   #"Output Barcode" := ("Expected/Value_All".V = "Expected/Value_All".Expected_1) OR ("Expected/Value_All".V = "Expected/Value_All".Expected_2) OR ("Expected/Value_All".V = "Expected/Value_All".Expected_3) OR ("Expected/Value_All".V = "Expected/Value_All".Expected_4) OR ("Expected/Value_All".V = "Expected/Value_All".Expected_5) OR ("Expected/Value_All".V = "Expected/Value_All".Expected_6) OR ("Expected/Value_All".V = "Expected/Value_All".Expected_7) OR ("Expected/Value_All".V = "Expected/Value_All".Expected_8) OR ("Expected/Value_All".V = "Expected/Value_All".Expected_9) OR ("Expected/Value_All".V = "Expected/Value_All".Expected_10) OR ("Expected/Value_All".V = "Expected/Value_All".Expected_11) OR ("Expected/Value_All".V = "Expected/Value_All".Expected_12) OR ("Expected/Value_All".V = "Expected/Value_All".Expected_13) OR ("Expected/Value_All".V = "Expected/Value_All".Expected_14) OR ("Expected/Value_All".V = "Expected/Value_All".Expected_15) OR ("Expected/Value_All".V = "Expected/Value_All".Expected_16) OR ("Expected/Value_All".V = "Expected/Value_All".Expected_17) OR ("Expected/Value_All".V = "Expected/Value_All".Expected_18) OR ("Expected/Value_All".V = "Expected/Value_All".Expected_19) OR ("Expected/Value_All".V = "Expected/Value_All".Expected_20) OR ("Expected/Value_All".V = "Expected/Value_All".Expected_21) OR ("Expected/Value_All".V = "Expected/Value_All".Expected_22) OR ("Expected/Value_All".V = "Expected/Value_All".Expected_23) OR ("Expected/Value_All".V = "Expected/Value_All".Expected_24) OR ("Expected/Value_All".V = "Expected/Value_All".Expected_25) OR ("Expected/Value_All".V = "Expected/Value_All".Expected_26) OR ("Expected/Value_All".V = "Expected/Value_All".Expected_27) OR ("Expected/Value_All".V = "Expected/Value_All".Expected_28) OR ("Expected/Value_All".V = "Expected/Value_All".Expected_29) OR ("Expected/Value_All".V = "Expected/Value_All".Expected_30) OR ("Expected/Value_All".V = "Expected/Value_All".Expected_31) OR ("Expected/Value_All".V = "Expected/Value_All".Expected_32) OR ("Expected/Value_All".V = "Expected/Value_All".Expected_33) OR ("Expected/Value_All".V = "Expected/Value_All".Expected_34) OR ("Expected/Value_All".V = "Expected/Value_All".Expected_35) OR ("Expected/Value_All".V = "Expected/Value_All".Expected_36) OR ("Expected/Value_All".V = "Expected/Value_All".Expected_37) OR ("Expected/Value_All".V = "Expected/Value_All".Expected_38) OR ("Expected/Value_All".V = "Expected/Value_All".Expected_39) OR ("Expected/Value_All".V = "Expected/Value_All".Expected_40) OR ("Expected/Value_All".V = "Expected/Value_All".Expected_41) OR ("Expected/Value_All".V = "Expected/Value_All".Expected_42) OR ("Expected/Value_All".V = "Expected/Value_All".Expected_43) OR ("Expected/Value_All".V = "Expected/Value_All".Expected_44) OR ("Expected/Value_All".V = "Expected/Value_All".Expected_45) OR ("Expected/Value_All".V = "Expected/Value_All".Expected_46) OR ("Expected/Value_All".V = "Expected/Value_All".Expected_47) OR ("Expected/Value_All".V = "Expected/Value_All".Expected_48) OR ("Expected/Value_All".V = "Expected/Value_All".Expected_49) OR ("Expected/Value_All".V = "Expected/Value_All".Expected_50) OR ("Expected/Value_All".V = "Expected/Value_All".Expected_51) OR ("Expected/Value_All".V = "Expected/Value_All".Expected_52) OR ("Expected/Value_All".V = "Expected/Value_All".Expected_53) OR ("Expected/Value_All".V = "Expected/Value_All".Expected_54) OR ("Expected/Value_All".V = "Expected/Value_All".Expected_55) OR ("Expected/Value_All".V = "Expected/Value_All".Expected_56) OR ("Expected/Value_All".V = "Expected/Value_All".Expected_57) OR ("Expected/Value_All".V = "Expected/Value_All".Expected_58) OR ("Expected/Value_All".V = "Expected/Value_All".Expected_59) OR ("Expected/Value_All".V = "Expected/Value_All".Expected_60) OR ("Expected/Value_All".V = "Expected/Value_All".Expected_61) OR ("Expected/Value_All".V = "Expected/Value_All".Expected_62) OR ("Expected/Value_All".V = "Expected/Value_All".Expected_63) OR ("Expected/Value_All".V = "Expected/Value_All".Expected_64) OR ("Expected/Value_All".V = "Expected/Value_All".Expected_65) OR ("Expected/Value_All".V = "Expected/Value_All".Expected_66) OR ("Expected/Value_All".V = "Expected/Value_All".Expected_67) OR ("Expected/Value_All".V = "Expected/Value_All".Expected_68) OR ("Expected/Value_All".V = "Expected/Value_All".Expected_69) OR ("Expected/Value_All".V = "Expected/Value_All".Expected_70) OR ("Expected/Value_All".V = "Expected/Value_All".Expected_71) OR ("Expected/Value_All".V = "Expected/Value_All".Expected_72) OR ("Expected/Value_All".V = "Expected/Value_All".Expected_73) OR ("Expected/Value_All".V = "Expected/Value_All".Expected_74) OR ("Expected/Value_All".V = "Expected/Value_All".Expected_75) OR ("Expected/Value_All".V = "Expected/Value_All".Expected_76) OR ("Expected/Value_All".V = "Expected/Value_All".Expected_77) OR ("Expected/Value_All".V = "Expected/Value_All".Expected_78) OR ("Expected/Value_All".V = "Expected/Value_All".Expected_79) OR ("Expected/Value_All".V = "Expected/Value_All".Expected_80) OR ("Expected/Value_All".V = "Expected/Value_All".Expected_81) OR ("Expected/Value_All".V = "Expected/Value_All".Expected_82) OR ("Expected/Value_All".V = "Expected/Value_All".Expected_83) OR ("Expected/Value_All".V = "Expected/Value_All".Expected_84) OR ("Expected/Value_All".V = "Expected/Value_All".Expected_85) OR ("Expected/Value_All".V = "Expected/Value_All".Expected_86) OR ("Expected/Value_All".V = "Expected/Value_All".Expected_87) OR ("Expected/Value_All".V = "Expected/Value_All".Expected_88) OR ("Expected/Value_All".V = "Expected/Value_All".Expected_89) OR ("Expected/Value_All".V = "Expected/Value_All".Expected_90) OR ("Expected/Value_All".V = "Expected/Value_All".Expected_91) OR ("Expected/Value_All".V = "Expected/Value_All".Expected_92) OR ("Expected/Value_All".V = "Expected/Value_All".Expected_93) OR ("Expected/Value_All".V = "Expected/Value_All".Expected_94) OR ("Expected/Value_All".V = "Expected/Value_All".Expected_95) OR ("Expected/Value_All".V = "Expected/Value_All".Expected_96) OR ("Expected/Value_All".V = "Expected/Value_All".Expected_97) OR ("Expected/Value_All".V = "Expected/Value_All".Expected_98) OR ("Expected/Value_All".V = "Expected/Value_All".Expected_99) OR ("Expected/Value_All".V = "Expected/Value_All".Expected_100) OR ("Expected/Value_All".V = "Expected/Value_All".Expected_101) OR ("Expected/Value_All".V = "Expected/Value_All".Expected_102) OR ("Expected/Value_All".V = "Expected/Value_All".Expected_103) OR ("Expected/Value_All".V = "Expected/Value_All".Expected_104) OR ("Expected/Value_All".V = "Expected/Value_All".Expected_105) OR ("Expected/Value_All".V = "Expected/Value_All".Expected_106) OR ("Expected/Value_All".V = "Expected/Value_All".Expected_107) OR ("Expected/Value_All".V = "Expected/Value_All".Expected_108) OR ("Expected/Value_All".V = "Expected/Value_All".Expected_109) OR ("Expected/Value_All".V = "Expected/Value_All".Expected_110) OR ("Expected/Value_All".V = "Expected/Value_All".Expected_111) OR ("Expected/Value_All".V = "Expected/Value_All".Expected_112) OR ("Expected/Value_All".V = "Expected/Value_All".Expected_113) OR ("Expected/Value_All".V = "Expected/Value_All".Expected_114) OR ("Expected/Value_All".V = "Expected/Value_All".Expected_115) OR ("Expected/Value_All".V = "Expected/Value_All".Expected_116) OR ("Expected/Value_All".V = "Expected/Value_All".Expected_117) OR ("Expected/Value_All".V = "Expected/Value_All".Expected_118) OR ("Expected/Value_All".V = "Expected/Value_All".Expected_119) OR ("Expected/Value_All".V = "Expected/Value_All".Expected_120) OR ("Expected/Value_All".V = "Expected/Value_All".Expected_121) OR ("Expected/Value_All".V = "Expected/Value_All".Expected_122) OR ("Expected/Value_All".V = "Expected/Value_All".Expected_123) OR ("Expected/Value_All".V = "Expected/Value_All".Expected_124) OR ("Expected/Value_All".V = "Expected/Value_All".Expected_125) OR ("Expected/Value_All".V = "Expected/Value_All".Expected_126) OR ("Expected/Value_All".V = "Expected/Value_All".Expected_127) OR ("Expected/Value_All".V = "Expected/Value_All".Expected_128) OR ("Expected/Value_All".V = "Expected/Value_All".Expected_129) OR ("Expected/Value_All".V = "Expected/Value_All".Expected_130) OR ("Expected/Value_All".V = "Expected/Value_All".Expected_131) OR ("Expected/Value_All".V = "Expected/Value_All".Expected_132) OR ("Expected/Value_All".V = "Expected/Value_All".Expected_133) OR ("Expected/Value_All".V = "Expected/Value_All".Expected_134) OR ("Expected/Value_All".V = "Expected/Value_All".Expected_135) OR ("Expected/Value_All".V = "Expected/Value_All".Expected_136) OR ("Expected/Value_All".V = "Expected/Value_All".Expected_137) OR ("Expected/Value_All".V = "Expected/Value_All".Expected_138) OR ("Expected/Value_All".V = "Expected/Value_All".Expected_139) OR ("Expected/Value_All".V = "Expected/Value_All".Expected_140) OR ("Expected/Value_All".V = "Expected/Value_All".Expected_141) OR ("Expected/Value_All".V = "Expected/Value_All".Expected_142) OR ("Expected/Value_All".V = "Expected/Value_All".Expected_143) OR ("Expected/Value_All".V = "Expected/Value_All".Expected_144) OR ("Expected/Value_All".V = "Expected/Value_All".Expected_145) OR ("Expected/Value_All".V = "Expected/Value_All".Expected_146) OR ("Expected/Value_All".V = "Expected/Value_All".Expected_147) OR ("Expected/Value_All".V = "Expected/Value_All".Expected_148) OR ("Expected/Value_All".V = "Expected/Value_All".Expected_149) OR ("Expected/Value_All".V = "Expected/Value_All".Expected_150) OR ("Expected/Value_All".V = "Expected/Value_All".Expected_151) OR ("Expected/Value_All".V = "Expected/Value_All".Expected_152) OR ("Expected/Value_All".V = "Expected/Value_All".Expected_153) OR ("Expected/Value_All".V = "Expected/Value_All".Expected_154) OR ("Expected/Value_All".V = "Expected/Value_All".Expected_155) OR ("Expected/Value_All".V = "Expected/Value_All".Expected_156) OR ("Expected/Value_All".V = "Expected/Value_All".Expected_157) OR ("Expected/Value_All".V = "Expected/Value_All".Expected_158) OR ("Expected/Value_All".V = "Expected/Value_All".Expected_159) OR ("Expected/Value_All".V = "Expected/Value_All".Expected_160) OR ("Expected/Value_All".V = "Expected/Value_All".Expected_161) OR ("Expected/Value_All".V = "Expected/Value_All".Expected_162) OR ("Expected/Value_All".V = "Expected/Value_All".Expected_163) OR ("Expected/Value_All".V = "Expected/Value_All".Expected_164) OR ("Expected/Value_All".V = "Expected/Value_All".Expected_165) OR ("Expected/Value_All".V = "Expected/Value_All".Expected_166) OR ("Expected/Value_All".V = "Expected/Value_All".Expected_167) OR ("Expected/Value_All".V = "Expected/Value_All".Expected_168) OR ("Expected/Value_All".V = "Expected/Value_All".Expected_169) OR ("Expected/Value_All".V = "Expected/Value_All".Expected_170) OR ("Expected/Value_All".V = "Expected/Value_All".Expected_171) OR ("Expected/Value_All".V = "Expected/Value_All".Expected_172) OR ("Expected/Value_All".V = "Expected/Value_All".Expected_173) OR ("Expected/Value_All".V = "Expected/Value_All".Expected_174) OR ("Expected/Value_All".V = "Expected/Value_All".Expected_175) OR ("Expected/Value_All".V = "Expected/Value_All".Expected_176) OR ("Expected/Value_All".V = "Expected/Value_All".Expected_177) OR ("Expected/Value_All".V = "Expected/Value_All".Expected_178) OR ("Expected/Value_All".V = "Expected/Value_All".Expected_179) OR ("Expected/Value_All".V = "Expected/Value_All".Expected_180) OR ("Expected/Value_All".V = "Expected/Value_All".Expected_181) OR ("Expected/Value_All".V = "Expected/Value_All".Expected_182) OR ("Expected/Value_All".V = "Expected/Value_All".Expected_183) OR ("Expected/Value_All".V = "Expected/Value_All".Expected_184) OR ("Expected/Value_All".V = "Expected/Value_All".Expected_185) OR ("Expected/Value_All".V = "Expected/Value_All".Expected_186) OR ("Expected/Value_All".V = "Expected/Value_All".Expected_187) OR ("Expected/Value_All".V = "Expected/Value_All".Expected_188) OR ("Expected/Value_All".V = "Expected/Value_All".Expected_189) OR ("Expected/Value_All".V = "Expected/Value_All".Expected_190) OR ("Expected/Value_All".V = "Expected/Value_All".Expected_191) OR ("Expected/Value_All".V = "Expected/Value_All".Expected_192) OR ("Expected/Value_All".V = "Expected/Value_All".Expected_193) OR ("Expected/Value_All".V = "Expected/Value_All".Expected_194) OR ("Expected/Value_All".V = "Expected/Value_All".Expected_195) OR ("Expected/Value_All".V = "Expected/Value_All".Expected_196) OR ("Expected/Value_All".V = "Expected/Value_All".Expected_197) OR ("Expected/Value_All".V = "Expected/Value_All".Expected_198) OR ("Expected/Value_All".V = "Expected/Value_All".Expected_199) OR ("Expected/Value_All".V = "Expected/Value_All".Expected_200) OR ("Expected/Value_All".V = "Expected/Value_All".Expected_201) OR ("Expected/Value_All".V = "Expected/Value_All".Expected_202) OR ("Expected/Value_All".V = "Expected/Value_All".Expected_203) OR ("Expected/Value_All".V = "Expected/Value_All".Expected_204) OR ("Expected/Value_All".V = "Expected/Value_All".Expected_205) OR ("Expected/Value_All".V = "Expected/Value_All".Expected_206) OR ("Expected/Value_All".V = "Expected/Value_All".Expected_207) OR ("Expected/Value_All".V = "Expected/Value_All".Expected_208) OR ("Expected/Value_All".V = "Expected/Value_All".Expected_209) OR ("Expected/Value_All".V = "Expected/Value_All".Expected_210) OR ("Expected/Value_All".V = "Expected/Value_All".Expected_211) OR ("Expected/Value_All".V = "Expected/Value_All".Expected_212) OR ("Expected/Value_All".V = "Expected/Value_All".Expected_213) OR ("Expected/Value_All".V = "Expected/Value_All".Expected_214) OR ("Expected/Value_All".V = "Expected/Value_All".Expected_215) OR ("Expected/Value_All".V = "Expected/Value_All".Expected_216) OR ("Expected/Value_All".V = "Expected/Value_All".Expected_217) OR ("Expected/Value_All".V = "Expected/Value_All".Expected_218) OR ("Expected/Value_All".V = "Expected/Value_All".Expected_219) OR ("Expected/Value_All".V = "Expected/Value_All".Expected_220) OR ("Expected/Value_All".V = "Expected/Value_All".Expected_221) OR ("Expected/Value_All".V = "Expected/Value_All".Expected_222) OR ("Expected/Value_All".V = "Expected/Value_All".Expected_223) OR ("Expected/Value_All".V = "Expected/Value_All".Expected_224) OR ("Expected/Value_All".V = "Expected/Value_All".Expected_225) OR ("Expected/Value_All".V = "Expected/Value_All".Expected_226) OR ("Expected/Value_All".V = "Expected/Value_All".Expected_227) OR ("Expected/Value_All".V = "Expected/Value_All".Expected_228) OR ("Expected/Value_All".V = "Expected/Value_All".Expected_229) OR ("Expected/Value_All".V = "Expected/Value_All".Expected_230) OR ("Expected/Value_All".V = "Expected/Value_All".Expected_231) OR ("Expected/Value_All".V = "Expected/Value_All".Expected_232) OR ("Expected/Value_All".V = "Expected/Value_All".Expected_233) OR ("Expected/Value_All".V = "Expected/Value_All".Expected_234) OR ("Expected/Value_All".V = "Expected/Value_All".Expected_235) OR ("Expected/Value_All".V = "Expected/Value_All".Expected_236) OR ("Expected/Value_All".V = "Expected/Value_All".Expected_237) OR ("Expected/Value_All".V = "Expected/Value_All".Expected_238) OR ("Expected/Value_All".V = "Expected/Value_All".Expected_239) OR ("Expected/Value_All".V = "Expected/Value_All".Expected_240) OR ("Expected/Value_All".V = "Expected/Value_All".Expected_241) OR ("Expected/Value_All".V = "Expected/Value_All".Expected_242) OR ("Expected/Value_All".V = "Expected/Value_All".Expected_243) OR ("Expected/Value_All".V = "Expected/Value_All".Expected_244) OR ("Expected/Value_All".V = "Expected/Value_All".Expected_245) OR ("Expected/Value_All".V = "Expected/Value_All".Expected_246) OR ("Expected/Value_All".V = "Expected/Value_All".Expected_247) OR ("Expected/Value_All".V = "Expected/Value_All".Expected_248) OR ("Expected/Value_All".V = "Expected/Value_All".Expected_249) OR ("Expected/Value_All".V = "Expected/Value_All".Expected_250) OR ("Expected/Value_All".V = "Expected/Value_All".Expected_251) OR ("Expected/Value_All".V = "Expected/Value_All".Expected_252) OR ("Expected/Value_All".V = "Expected/Value_All".Expected_253) OR ("Expected/Value_All".V = "Expected/Value_All".Expected_254) OR ("Expected/Value_All".V = "Expected/Value_All".Expected_255) OR ("Expected/Value_All".V = "Expected/Value_All".Expected_256) OR ("Expected/Value_All".V = "Expected/Value_All".Expected_257) OR ("Expected/Value_All".V = "Expected/Value_All".Expected_258) OR ("Expected/Value_All".V = "Expected/Value_All".Expected_259) OR ("Expected/Value_All".V = "Expected/Value_All".Expected_260) OR ("Expected/Value_All".V = "Expected/Value_All".Expected_261) OR ("Expected/Value_All".V = "Expected/Value_All".Expected_262) OR ("Expected/Value_All".V = "Expected/Value_All".Expected_263) OR ("Expected/Value_All".V = "Expected/Value_All".Expected_264) OR ("Expected/Value_All".V = "Expected/Value_All".Expected_265) OR ("Expected/Value_All".V = "Expected/Value_All".Expected_266) OR ("Expected/Value_All".V = "Expected/Value_All".Expected_267) OR ("Expected/Value_All".V = "Expected/Value_All".Expected_268) OR ("Expected/Value_All".V = "Expected/Value_All".Expected_269) OR ("Expected/Value_All".V = "Expected/Value_All".Expected_270) OR ("Expected/Value_All".V = "Expected/Value_All".Expected_271) OR ("Expected/Value_All".V = "Expected/Value_All".Expected_272) OR ("Expected/Value_All".V = "Expected/Value_All".Expected_273) OR ("Expected/Value_All".V = "Expected/Value_All".Expected_274) OR ("Expected/Value_All".V = "Expected/Value_All".Expected_275) OR ("Expected/Value_All".V = "Expected/Value_All".Expected_276) OR ("Expected/Value_All".V = "Expected/Value_All".Expected_277) OR ("Expected/Value_All".V = "Expected/Value_All".Expected_278) OR ("Expected/Value_All".V = "Expected/Value_All".Expected_279) OR ("Expected/Value_All".V = "Expected/Value_All".Expected_280) OR ("Expected/Value_All".V = "Expected/Value_All".Expected_281) OR ("Expected/Value_All".V = "Expected/Value_All".Expected_282) OR ("Expected/Value_All".V = "Expected/Value_All".Expected_283) OR ("Expected/Value_All".V = "Expected/Value_All".Expected_284) OR ("Expected/Value_All".V = "Expected/Value_All".Expected_285) OR ("Expected/Value_All".V = "Expected/Value_All".Expected_286) OR ("Expected/Value_All".V = "Expected/Value_All".Expected_287) OR ("Expected/Value_All".V = "Expected/Value_All".Expected_288) OR ("Expected/Value_All".V = "Expected/Value_All".Expected_289) OR ("Expected/Value_All".V = "Expected/Value_All".Expected_290) OR ("Expected/Value_All".V = "Expected/Value_All".Expected_291) OR ("Expected/Value_All".V = "Expected/Value_All".Expected_292) OR ("Expected/Value_All".V = "Expected/Value_All".Expected_293) OR ("Expected/Value_All".V = "Expected/Value_All".Expected_294) OR ("Expected/Value_All".V = "Expected/Value_All".Expected_295) OR ("Expected/Value_All".V = "Expected/Value_All".Expected_296) OR ("Expected/Value_All".V = "Expected/Value_All".Expected_297) OR ("Expected/Value_All".V = "Expected/Value_All".Expected_298) OR ("Expected/Value_All".V = "Expected/Value_All".Expected_299) OR ("Expected/Value_All".V = "Expected/Value_All".Expected_300) OR ("Expected/Value_All".V = "Expected/Value_All".Expected_301) OR ("Expected/Value_All".V = "Expected/Value_All".Expected_302) OR ("Expected/Value_All".V = "Expected/Value_All".Expected_303) OR ("Expected/Value_All".V = "Expected/Value_All".Expected_304) OR ("Expected/Value_All".V = "Expected/Value_All".Expected_305) OR ("Expected/Value_All".V = "Expected/Value_All".Expected_306) OR ("Expected/Value_All".V = "Expected/Value_All".Expected_307) OR ("Expected/Value_All".V = "Expected/Value_All".Expected_308) OR ("Expected/Value_All".V = "Expected/Value_All".Expected_309) OR ("Expected/Value_All".V = "Expected/Value_All".Expected_310) OR ("Expected/Value_All".V = "Expected/Value_All".Expected_311) OR ("Expected/Value_All".V = "Expected/Value_All".Expected_312) OR ("Expected/Value_All".V = "Expected/Value_All".Expected_313) OR ("Expected/Value_All".V = "Expected/Value_All".Expected_314) OR ("Expected/Value_All".V = "Expected/Value_All".Expected_315) OR ("Expected/Value_All".V = "Expected/Value_All".Expected_316) OR ("Expected/Value_All".V = "Expected/Value_All".Expected_317) OR ("Expected/Value_All".V = "Expected/Value_All".Expected_318) OR ("Expected/Value_All".V = "Expected/Value_All".Expected_319) OR ("Expected/Value_All".V = "Expected/Value_All".Expected_320) OR ("Expected/Value_All".V = "Expected/Value_All".Expected_321) OR ("Expected/Value_All".V = "Expected/Value_All".Expected_322) OR ("Expected/Value_All".V = "Expected/Value_All".Expected_323) OR ("Expected/Value_All".V = "Expected/Value_All".Expected_324) OR ("Expected/Value_All".V = "Expected/Value_All".Expected_325) OR ("Expected/Value_All".V = "Expected/Value_All".Expected_326) OR ("Expected/Value_All".V = "Expected/Value_All".Expected_327) OR ("Expected/Value_All".V = "Expected/Value_All".Expected_328) OR ("Expected/Value_All".V = "Expected/Value_All".Expected_329) OR ("Expected/Value_All".V = "Expected/Value_All".Expected_330) OR ("Expected/Value_All".V = "Expected/Value_All".Expected_331) OR ("Expected/Value_All".V = "Expected/Value_All".Expected_332) OR ("Expected/Value_All".V = "Expected/Value_All".Expected_333) OR ("Expected/Value_All".V = "Expected/Value_All".Expected_334) OR ("Expected/Value_All".V = "Expected/Value_All".Expected_335) OR ("Expected/Value_All".V = "Expected/Value_All".Expected_336) OR ("Expected/Value_All".V = "Expected/Value_All".Expected_337) OR ("Expected/Value_All".V = "Expected/Value_All".Expected_338) OR ("Expected/Value_All".V = "Expected/Value_All".Expected_339) OR ("Expected/Value_All".V = "Expected/Value_All".Expected_340) OR ("Expected/Value_All".V = "Expected/Value_All".Expected_341) OR ("Expected/Value_All".V = "Expected/Value_All".Expected_342) OR ("Expected/Value_All".V = "Expected/Value_All".Expected_343) OR ("Expected/Value_All".V = "Expected/Value_All".Expected_344) OR ("Expected/Value_All".V = "Expected/Value_All".Expected_345) OR ("Expected/Value_All".V = "Expected/Value_All".Expected_346) OR ("Expected/Value_All".V = "Expected/Value_All".Expected_347) OR ("Expected/Value_All".V = "Expected/Value_All".Expected_348) OR ("Expected/Value_All".V = "Expected/Value_All".Expected_349) OR ("Expected/Value_All".V = "Expected/Value_All".Expected_350) OR ("Expected/Value_All".V = "Expected/Value_All".Expected_351) OR ("Expected/Value_All".V = "Expected/Value_All".Expected_352) OR ("Expected/Value_All".V = "Expected/Value_All".Expected_353) OR ("Expected/Value_All".V = "Expected/Value_All".Expected_354) OR ("Expected/Value_All".V = "Expected/Value_All".Expected_355) OR ("Expected/Value_All".V = "Expected/Value_All".Expected_356) OR ("Expected/Value_All".V = "Expected/Value_All".Expected_357) OR ("Expected/Value_All".V = "Expected/Value_All".Expected_358) OR ("Expected/Value_All".V = "Expected/Value_All".Expected_359) OR ("Expected/Value_All".V = "Expected/Value_All".Expected_360) OR ("Expected/Value_All".V = "Expected/Value_All".Expected_361) OR ("Expected/Value_All".V = "Expected/Value_All".Expected_362) OR ("Expected/Value_All".V = "Expected/Value_All".Expected_363) OR ("Expected/Value_All".V = "Expected/Value_All".Expected_364) OR ("Expected/Value_All".V = "Expected/Value_All".Expected_365) OR ("Expected/Value_All".V = "Expected/Value_All".Expected_366) OR ("Expected/Value_All".V = "Expected/Value_All".Expected_367) OR ("Expected/Value_All".V = "Expected/Value_All".Expected_368) OR ("Expected/Value_All".V = "Expected/Value_All".Expected_369) OR ("Expected/Value_All".V = "Expected/Value_All".Expected_370) OR ("Expected/Value_All".V = "Expected/Value_All".Expected_371) OR ("Expected/Value_All".V = "Expected/Value_All".Expected_372) OR ("Expected/Value_All".V = "Expected/Value_All".Expected_373) OR ("Expected/Value_All".V = "Expected/Value_All".Expected_374) OR ("Expected/Value_All".V = "Expected/Value_All".Expected_375) OR ("Expected/Value_All".V = "Expected/Value_All".Expected_376) OR ("Expected/Value_All".V = "Expected/Value_All".Expected_377) OR ("Expected/Value_All".V = "Expected/Value_All".Expected_378) OR ("Expected/Value_All".V = "Expected/Value_All".Expected_379) OR ("Expected/Value_All".V = "Expected/Value_All".Expected_380) OR ("Expected/Value_All".V = "Expected/Value_All".Expected_381) OR ("Expected/Value_All".V = "Expected/Value_All".Expected_382) OR ("Expected/Value_All".V = "Expected/Value_All".Expected_383) OR ("Expected/Value_All".V = "Expected/Value_All".Expected_384) OR ("Expected/Value_All".V = "Expected/Value_All".Expected_385) OR ("Expected/Value_All".V = "Expected/Value_All".Expected_386) OR ("Expected/Value_All".V = "Expected/Value_All".Expected_387) OR ("Expected/Value_All".V = "Expected/Value_All".Expected_388) OR ("Expected/Value_All".V = "Expected/Value_All".Expected_389) OR ("Expected/Value_All".V = "Expected/Value_All".Expected_390) OR ("Expected/Value_All".V = "Expected/Value_All".Expected_391) OR ("Expected/Value_All".V = "Expected/Value_All".Expected_392) OR ("Expected/Value_All".V = "Expected/Value_All".Expected_393) OR ("Expected/Value_All".V = "Expected/Value_All".Expected_394) OR ("Expected/Value_All".V = "Expected/Value_All".Expected_395) OR ("Expected/Value_All".V = "Expected/Value_All".Expected_396) OR ("Expected/Value_All".V = "Expected/Value_All".Expected_397) OR ("Expected/Value_All".V = "Expected/Value_All".Expected_398) OR ("Expected/Value_All".V = "Expected/Value_All".Expected_399) OR ("Expected/Value_All".V = "Expected/Value_All".Expected_400) OR ("Expected/Value_All".V = "Expected/Value_All".Expected_401) OR ("Expected/Value_All".V = "Expected/Value_All".Expected_402) OR ("Expected/Value_All".V = "Expected/Value_All".Expected_403) OR ("Expected/Value_All".V = "Expected/Value_All".Expected_404) OR ("Expected/Value_All".V = "Expected/Value_All".Expected_405) OR ("Expected/Value_All".V = "Expected/Value_All".Expected_406) OR ("Expected/Value_All".V = "Expected/Value_All".Expected_407) OR ("Expected/Value_All".V = "Expected/Value_All".Expected_408) OR ("Expected/Value_All".V = "Expected/Value_All".Expected_409) OR ("Expected/Value_All".V = "Expected/Value_All".Expected_410) OR ("Expected/Value_All".V = "Expected/Value_All".Expected_411) OR ("Expected/Value_All".V = "Expected/Value_All".Expected_412) OR ("Expected/Value_All".V = "Expected/Value_All".Expected_413) OR ("Expected/Value_All".V = "Expected/Value_All".Expected_414) OR ("Expected/Value_All".V = "Expected/Value_All".Expected_415) OR ("Expected/Value_All".V = "Expected/Value_All".Expected_416) OR ("Expected/Value_All".V = "Expected/Value_All".Expected_417) OR ("Expected/Value_All".V = "Expected/Value_All".Expected_418) OR ("Expected/Value_All".V = "Expected/Value_All".Expected_419) OR ("Expected/Value_All".V = "Expected/Value_All".Expected_420) OR ("Expected/Value_All".V = "Expected/Value_All".Expected_421) OR ("Expected/Value_All".V = "Expected/Value_All".Expected_422) OR ("Expected/Value_All".V = "Expected/Value_All".Expected_423) OR ("Expected/Value_All".V = "Expected/Value_All".Expected_424) OR ("Expected/Value_All".V = "Expected/Value_All".Expected_425) OR ("Expected/Value_All".V = "Expected/Value_All".Expected_426) OR ("Expected/Value_All".V = "Expected/Value_All".Expected_427) OR ("Expected/Value_All".V = "Expected/Value_All".Expected_428) OR ("Expected/Value_All".V = "Expected/Value_All".Expected_429) OR ("Expected/Value_All".V = "Expected/Value_All".Expected_430) OR ("Expected/Value_All".V = "Expected/Value_All".Expected_431) OR ("Expected/Value_All".V = "Expected/Value_All".Expected_432) OR ("Expected/Value_All".V = "Expected/Value_All".Expected_433) OR ("Expected/Value_All".V = "Expected/Value_All".Expected_434) OR ("Expected/Value_All".V = "Expected/Value_All".Expected_435) OR ("Expected/Value_All".V = "Expected/Value_All".Expected_436) OR ("Expected/Value_All".V = "Expected/Value_All".Expected_437) OR ("Expected/Value_All".V = "Expected/Value_All".Expected_438) OR ("Expected/Value_All".V = "Expected/Value_All".Expected_439) OR ("Expected/Value_All".V = "Expected/Value_All".Expected_440) OR ("Expected/Value_All".V = "Expected/Value_All".Expected_441) OR ("Expected/Value_All".V = "Expected/Value_All".Expected_442) OR ("Expected/Value_All".V = "Expected/Value_All".Expected_443) OR ("Expected/Value_All".V = "Expected/Value_All".Expected_444) OR ("Expected/Value_All".V = "Expected/Value_All".Expected_445) OR ("Expected/Value_All".V = "Expected/Value_All".Expected_446) OR ("Expected/Value_All".V = "Expected/Value_All".Expected_447) OR ("Expected/Value_All".V = "Expected/Value_All".Expected_448) OR ("Expected/Value_All".V = "Expected/Value_All".Expected_449) OR ("Expected/Value_All".V = "Expected/Value_All".Expected_450) OR ("Expected/Value_All".V = "Expected/Value_All".Expected_451) OR ("Expected/Value_All".V = "Expected/Value_All".Expected_452) OR ("Expected/Value_All".V = "Expected/Value_All".Expected_453) OR ("Expected/Value_All".V = "Expected/Value_All".Expected_454) OR ("Expected/Value_All".V = "Expected/Value_All".Expected_455) OR ("Expected/Value_All".V = "Expected/Value_All".Expected_456) OR ("Expected/Value_All".V = "Expected/Value_All".Expected_457) OR ("Expected/Value_All".V = "Expected/Value_All".Expected_458) OR ("Expected/Value_All".V = "Expected/Value_All".Expected_459) OR ("Expected/Value_All".V = "Expected/Value_All".Expected_460) OR ("Expected/Value_All".V = "Expected/Value_All".Expected_461) OR ("Expected/Value_All".V = "Expected/Value_All".Expected_462) OR ("Expected/Value_All".V = "Expected/Value_All".Expected_463) OR ("Expected/Value_All".V = "Expected/Value_All".Expected_464) OR ("Expected/Value_All".V = "Expected/Value_All".Expected_465) OR ("Expected/Value_All".V = "Expected/Value_All".Expected_466) OR ("Expected/Value_All".V = "Expected/Value_All".Expected_467) OR ("Expected/Value_All".V = "Expected/Value_All".Expected_468) OR ("Expected/Value_All".V = "Expected/Value_All".Expected_469) OR ("Expected/Value_All".V = "Expected/Value_All".Expected_470) OR ("Expected/Value_All".V = "Expected/Value_All".Expected_471) OR ("Expected/Value_All".V = "Expected/Value_All".Expected_472) OR ("Expected/Value_All".V = "Expected/Value_All".Expected_473) OR ("Expected/Value_All".V = "Expected/Value_All".Expected_474) OR ("Expected/Value_All".V = "Expected/Value_All".Expected_475) OR ("Expected/Value_All".V = "Expected/Value_All".Expected_476) OR ("Expected/Value_All".V = "Expected/Value_All".Expected_477) OR ("Expected/Value_All".V = "Expected/Value_All".Expected_478) OR ("Expected/Value_All".V = "Expected/Value_All".Expected_479) OR ("Expected/Value_All".V = "Expected/Value_All".Expected_480) OR ("Expected/Value_All".V = "Expected/Value_All".Expected_481) OR ("Expected/Value_All".V = "Expected/Value_All".Expected_482) OR ("Expected/Value_All".V = "Expected/Value_All".Expected_483) OR ("Expected/Value_All".V = "Expected/Value_All".Expected_484) OR ("Expected/Value_All".V = "Expected/Value_All".Expected_485) OR ("Expected/Value_All".V = "Expected/Value_All".Expected_486) OR ("Expected/Value_All".V = "Expected/Value_All".Expected_487) OR ("Expected/Value_All".V = "Expected/Value_All".Expected_488) OR ("Expected/Value_All".V = "Expected/Value_All".Expected_489) OR ("Expected/Value_All".V = "Expected/Value_All".Expected_490) OR ("Expected/Value_All".V = "Expected/Value_All".Expected_491) OR ("Expected/Value_All".V = "Expected/Value_All".Expected_492) OR ("Expected/Value_All".V = "Expected/Value_All".Expected_493) OR ("Expected/Value_All".V = "Expected/Value_All".Expected_494) OR ("Expected/Value_All".V = "Expected/Value_All".Expected_495) OR ("Expected/Value_All".V = "Expected/Value_All".Expected_496) OR ("Expected/Value_All".V = "Expected/Value_All".Expected_497) OR ("Expected/Value_All".V = "Expected/Value_All".Expected_498) OR ("Expected/Value_All".V = "Expected/Value_All".Expected_499) OR ("Expected/Value_All".V = "Expected/Value_All".Expected_500) OR ("Expected/Value_All".V = "Expected/Value_All".Expected_501) OR ("Expected/Value_All".V = "Expected/Value_All".Expected_502) OR ("Expected/Value_All".V = "Expected/Value_All".Expected_503) OR ("Expected/Value_All".V = "Expected/Value_All".Expected_504) OR ("Expected/Value_All".V = "Expected/Value_All".Expected_505) OR ("Expected/Value_All".V = "Expected/Value_All".Expected_506) OR ("Expected/Value_All".V = "Expected/Value_All".Expected_507) OR ("Expected/Value_All".V = "Expected/Value_All".Expected_508) OR ("Expected/Value_All".V = "Expected/Value_All".Expected_509) OR ("Expected/Value_All".V = "Expected/Value_All".Expected_510) OR ("Expected/Value_All".V = "Expected/Value_All".Expected_511) OR ("Expected/Value_All".V = "Expected/Value_All".Expected_512) OR ("Expected/Value_All".V = "Expected/Value_All".Expected_513) OR ("Expected/Value_All".V = "Expected/Value_All".Expected_514) OR ("Expected/Value_All".V = "Expected/Value_All".Expected_515) OR ("Expected/Value_All".V = "Expected/Value_All".Expected_516) OR ("Expected/Value_All".V = "Expected/Value_All".Expected_517) OR ("Expected/Value_All".V = "Expected/Value_All".Expected_518) OR ("Expected/Value_All".V = "Expected/Value_All".Expected_519) OR ("Expected/Value_All".V = "Expected/Value_All".Expected_520);
END_REGION
END_FUNCTION

FUNCTION "Expected" : Void   // FC3, LAD
{ S7_Optimized_Access := 'TRUE' }
VERSION : 0.1
   VAR_INPUT
      Expected1 : String;
      Expected2 : String;
      Expected3 : String;
      Expected4 : String;
      Expected5 : String;
      Expected6 : String;
      Expected7 : String;
      Expected8 : String;
      Expected9 : String;
      Expected10 : String;
      Expected11 : String;
      Expected12 : String;
      Expected13 : String;
      Expected14 : String;
      Expected15 : String;
      Expected16 : String;
      Expected17 : String;
      Expected18 : String;
      Expected19 : String;
      Expected20 : String;
      Expected21 : String;
      Expected22 : String;
      Expected23 : String;
      Expected24 : String;
      Expected25 : String;
      Expected26 : String;
   END_VAR
   VAR_OUTPUT
      On_Motor : Bool;
   END_VAR
BEGIN

REGION Network 1
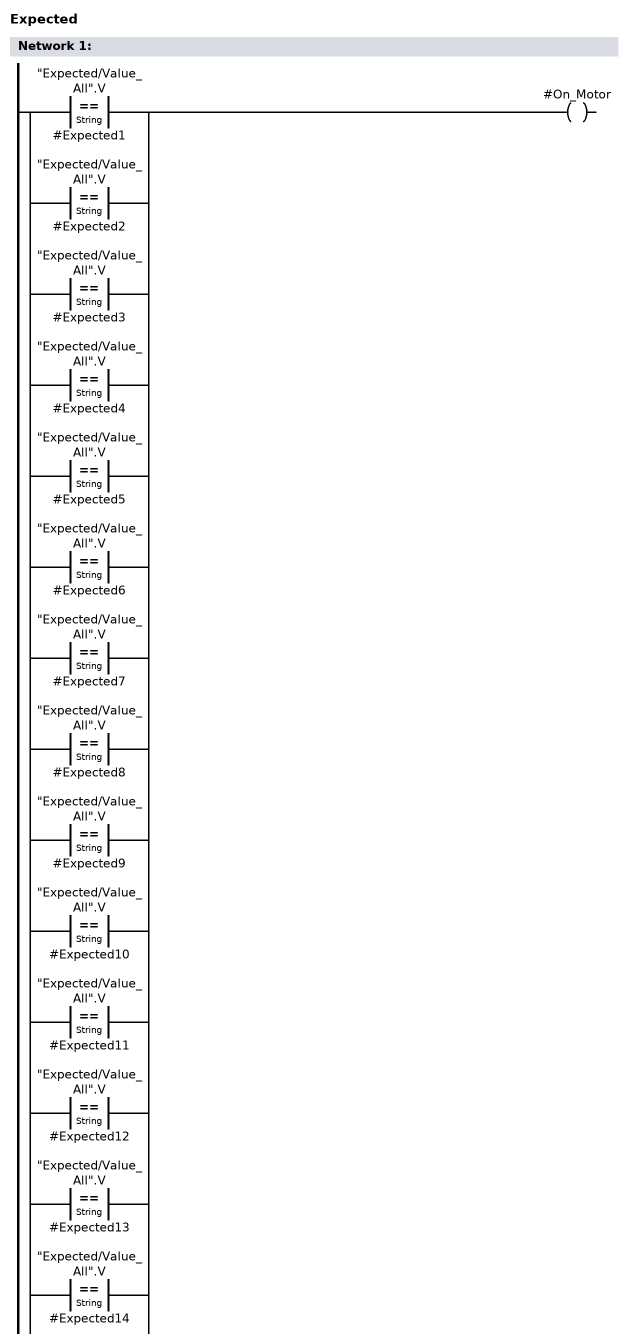
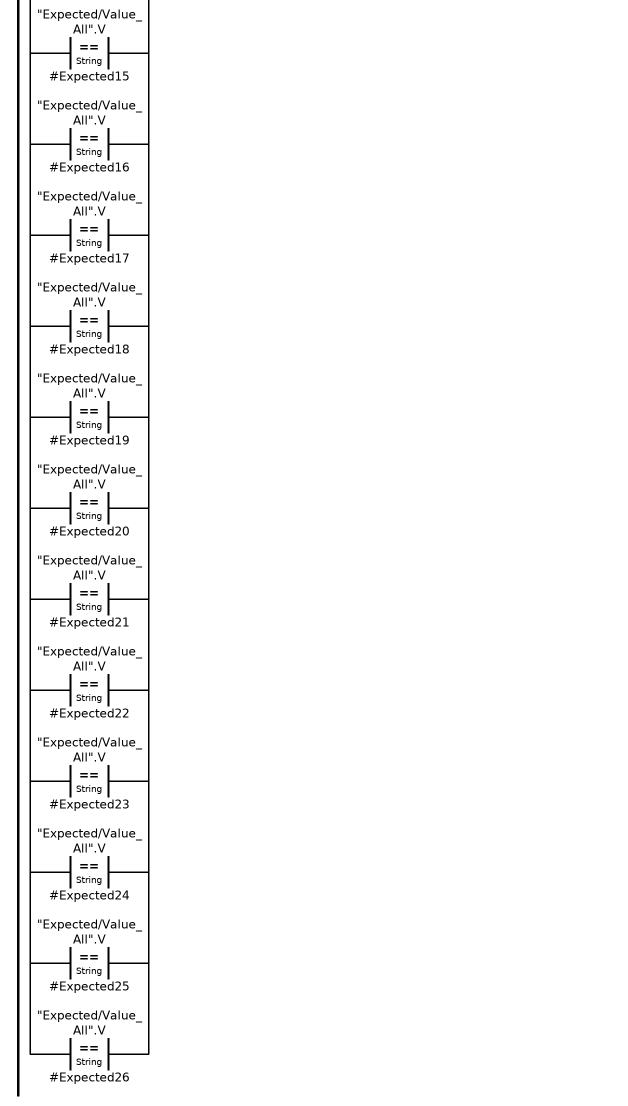
   RUNG wire#powerrail
      { S7_Templates := "SrcType := String" } EQ_Contact(in1 := "Expected/Value_All".V, in2 := #Expected1)
      wire#w1
      Coil( #On_Motor )
   END_RUNG
   RUNG wire#powerrail
      { S7_Templates := "SrcType := String" } EQ_Contact(in1 := "Expected/Value_All".V, in2 := #Expected2)
   END_RUNG wire#w1
   RUNG wire#powerrail
      { S7_Templates := "SrcType := String" } EQ_Contact(in1 := "Expected/Value_All".V, in2 := #Expected3)
   END_RUNG wire#w1
   RUNG wire#powerrail
      { S7_Templates := "SrcType := String" } EQ_Contact(in1 := "Expected/Value_All".V, in2 := #Expected4)
   END_RUNG wire#w1
   RUNG wire#powerrail
      { S7_Templates := "SrcType := String" } EQ_Contact(in1 := "Expected/Value_All".V, in2 := #Expected5)
   END_RUNG wire#w1
   RUNG wire#powerrail
      { S7_Templates := "SrcType := String" } EQ_Contact(in1 := "Expected/Value_All".V, in2 := #Expected6)
   END_RUNG wire#w1
   RUNG wire#powerrail
      { S7_Templates := "SrcType := String" } EQ_Contact(in1 := "Expected/Value_All".V, in2 := #Expected7)
   END_RUNG wire#w1
   RUNG wire#powerrail
      { S7_Templates := "SrcType := String" } EQ_Contact(in1 := "Expected/Value_All".V, in2 := #Expected8)
   END_RUNG wire#w1
   RUNG wire#powerrail
      { S7_Templates := "SrcType := String" } EQ_Contact(in1 := "Expected/Value_All".V, in2 := #Expected9)
   END_RUNG wire#w1
   RUNG wire#powerrail
      { S7_Templates := "SrcType := String" } EQ_Contact(in1 := "Expected/Value_All".V, in2 := #Expected10)
   END_RUNG wire#w1
   RUNG wire#powerrail
      { S7_Templates := "SrcType := String" } EQ_Contact(in1 := "Expected/Value_All".V, in2 := #Expected11)
   END_RUNG wire#w1
   RUNG wire#powerrail
      { S7_Templates := "SrcType := String" } EQ_Contact(in1 := "Expected/Value_All".V, in2 := #Expected12)
   END_RUNG wire#w1
   RUNG wire#powerrail
      { S7_Templates := "SrcType := String" } EQ_Contact(in1 := "Expected/Value_All".V, in2 := #Expected13)
   END_RUNG wire#w1
   RUNG wire#powerrail
      { S7_Templates := "SrcType := String" } EQ_Contact(in1 := "Expected/Value_All".V, in2 := #Expected14)
   END_RUNG wire#w1
   RUNG wire#powerrail
      { S7_Templates := "SrcType := String" } EQ_Contact(in1 := "Expected/Value_All".V, in2 := #Expected15)
   END_RUNG wire#w1
   RUNG wire#powerrail
      { S7_Templates := "SrcType := String" } EQ_Contact(in1 := "Expected/Value_All".V, in2 := #Expected16)
   END_RUNG wire#w1
   RUNG wire#powerrail
      { S7_Templates := "SrcType := String" } EQ_Contact(in1 := "Expected/Value_All".V, in2 := #Expected17)
   END_RUNG wire#w1
   RUNG wire#powerrail
      { S7_Templates := "SrcType := String" } EQ_Contact(in1 := "Expected/Value_All".V, in2 := #Expected18)
   END_RUNG wire#w1
   RUNG wire#powerrail
      { S7_Templates := "SrcType := String" } EQ_Contact(in1 := "Expected/Value_All".V, in2 := #Expected19)
   END_RUNG wire#w1
   RUNG wire#powerrail
      { S7_Templates := "SrcType := String" } EQ_Contact(in1 := "Expected/Value_All".V, in2 := #Expected20)
   END_RUNG wire#w1
   RUNG wire#powerrail
      { S7_Templates := "SrcType := String" } EQ_Contact(in1 := "Expected/Value_All".V, in2 := #Expected21)
   END_RUNG wire#w1
   RUNG wire#powerrail
      { S7_Templates := "SrcType := String" } EQ_Contact(in1 := "Expected/Value_All".V, in2 := #Expected22)
   END_RUNG wire#w1
   RUNG wire#powerrail
      { S7_Templates := "SrcType := String" } EQ_Contact(in1 := "Expected/Value_All".V, in2 := #Expected23)
   END_RUNG wire#w1
   RUNG wire#powerrail
      { S7_Templates := "SrcType := String" } EQ_Contact(in1 := "Expected/Value_All".V, in2 := #Expected24)
   END_RUNG wire#w1
   RUNG wire#powerrail
      { S7_Templates := "SrcType := String" } EQ_Contact(in1 := "Expected/Value_All".V, in2 := #Expected25)
   END_RUNG wire#w1
   RUNG wire#powerrail
      { S7_Templates := "SrcType := String" } EQ_Contact(in1 := "Expected/Value_All".V, in2 := #Expected26)
   END_RUNG wire#w1
   // the same network as SCL:
   #On_Motor := ("Expected/Value_All".V = #Expected1) OR ("Expected/Value_All".V = #Expected2) OR ("Expected/Value_All".V = #Expected3) OR ("Expected/Value_All".V = #Expected4) OR ("Expected/Value_All".V = #Expected5) OR ("Expected/Value_All".V = #Expected6) OR ("Expected/Value_All".V = #Expected7) OR ("Expected/Value_All".V = #Expected8) OR ("Expected/Value_All".V = #Expected9) OR ("Expected/Value_All".V = #Expected10) OR ("Expected/Value_All".V = #Expected11) OR ("Expected/Value_All".V = #Expected12) OR ("Expected/Value_All".V = #Expected13) OR ("Expected/Value_All".V = #Expected14) OR ("Expected/Value_All".V = #Expected15) OR ("Expected/Value_All".V = #Expected16) OR ("Expected/Value_All".V = #Expected17) OR ("Expected/Value_All".V = #Expected18) OR ("Expected/Value_All".V = #Expected19) OR ("Expected/Value_All".V = #Expected20) OR ("Expected/Value_All".V = #Expected21) OR ("Expected/Value_All".V = #Expected22) OR ("Expected/Value_All".V = #Expected23) OR ("Expected/Value_All".V = #Expected24) OR ("Expected/Value_All".V = #Expected25) OR ("Expected/Value_All".V = #Expected26);
END_REGION
END_FUNCTION

FUNCTION "Ex(20ช่อง)" : Void   // FC4, LAD
{ S7_Optimized_Access := 'TRUE' }
VERSION : 0.1
   VAR_INPUT
      Expected1 : String;
      Expected2 : String;
      Expected3 : String;
      Expected4 : String;
      Expected5 : String;
      Expected6 : String;
      Expected7 : String;
      Expected8 : String;
      Expected9 : String;
      Expected10 : String;
      Expected11 : String;
      Expected12 : String;
      Expected13 : String;
      Expected14 : String;
      Expected15 : String;
      Expected16 : String;
      Expected17 : String;
      Expected18 : String;
      Expected19 : String;
      Expected20 : String;
   END_VAR
   VAR_OUTPUT
      On_Motor : Bool;
   END_VAR
BEGIN

REGION Network 1
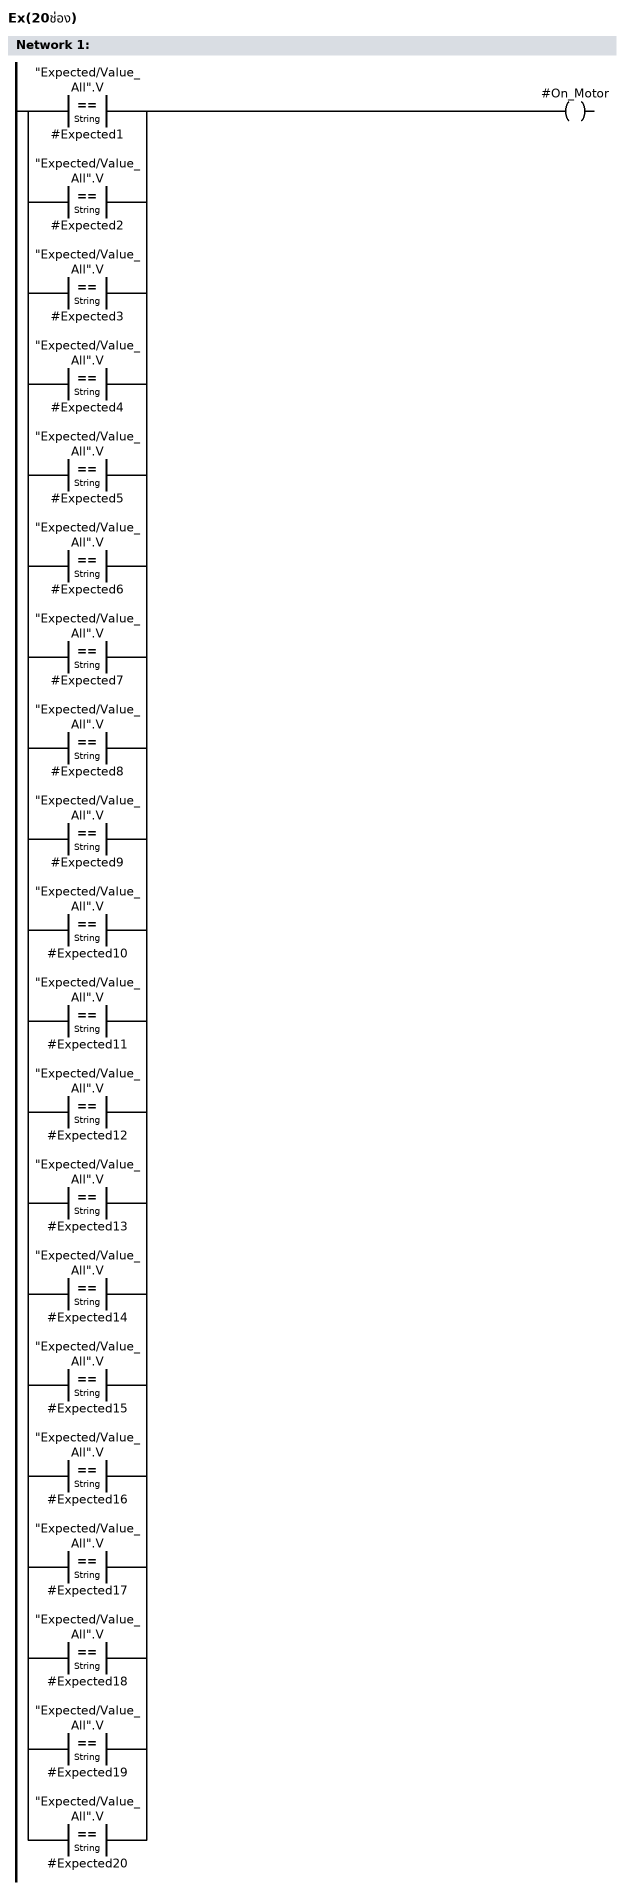
   RUNG wire#powerrail
      { S7_Templates := "SrcType := String" } EQ_Contact(in1 := "Expected/Value_All".V, in2 := #Expected1)
      wire#w1
      Coil( #On_Motor )
   END_RUNG
   RUNG wire#powerrail
      { S7_Templates := "SrcType := String" } EQ_Contact(in1 := "Expected/Value_All".V, in2 := #Expected2)
   END_RUNG wire#w1
   RUNG wire#powerrail
      { S7_Templates := "SrcType := String" } EQ_Contact(in1 := "Expected/Value_All".V, in2 := #Expected3)
   END_RUNG wire#w1
   RUNG wire#powerrail
      { S7_Templates := "SrcType := String" } EQ_Contact(in1 := "Expected/Value_All".V, in2 := #Expected4)
   END_RUNG wire#w1
   RUNG wire#powerrail
      { S7_Templates := "SrcType := String" } EQ_Contact(in1 := "Expected/Value_All".V, in2 := #Expected5)
   END_RUNG wire#w1
   RUNG wire#powerrail
      { S7_Templates := "SrcType := String" } EQ_Contact(in1 := "Expected/Value_All".V, in2 := #Expected6)
   END_RUNG wire#w1
   RUNG wire#powerrail
      { S7_Templates := "SrcType := String" } EQ_Contact(in1 := "Expected/Value_All".V, in2 := #Expected7)
   END_RUNG wire#w1
   RUNG wire#powerrail
      { S7_Templates := "SrcType := String" } EQ_Contact(in1 := "Expected/Value_All".V, in2 := #Expected8)
   END_RUNG wire#w1
   RUNG wire#powerrail
      { S7_Templates := "SrcType := String" } EQ_Contact(in1 := "Expected/Value_All".V, in2 := #Expected9)
   END_RUNG wire#w1
   RUNG wire#powerrail
      { S7_Templates := "SrcType := String" } EQ_Contact(in1 := "Expected/Value_All".V, in2 := #Expected10)
   END_RUNG wire#w1
   RUNG wire#powerrail
      { S7_Templates := "SrcType := String" } EQ_Contact(in1 := "Expected/Value_All".V, in2 := #Expected11)
   END_RUNG wire#w1
   RUNG wire#powerrail
      { S7_Templates := "SrcType := String" } EQ_Contact(in1 := "Expected/Value_All".V, in2 := #Expected12)
   END_RUNG wire#w1
   RUNG wire#powerrail
      { S7_Templates := "SrcType := String" } EQ_Contact(in1 := "Expected/Value_All".V, in2 := #Expected13)
   END_RUNG wire#w1
   RUNG wire#powerrail
      { S7_Templates := "SrcType := String" } EQ_Contact(in1 := "Expected/Value_All".V, in2 := #Expected14)
   END_RUNG wire#w1
   RUNG wire#powerrail
      { S7_Templates := "SrcType := String" } EQ_Contact(in1 := "Expected/Value_All".V, in2 := #Expected15)
   END_RUNG wire#w1
   RUNG wire#powerrail
      { S7_Templates := "SrcType := String" } EQ_Contact(in1 := "Expected/Value_All".V, in2 := #Expected16)
   END_RUNG wire#w1
   RUNG wire#powerrail
      { S7_Templates := "SrcType := String" } EQ_Contact(in1 := "Expected/Value_All".V, in2 := #Expected17)
   END_RUNG wire#w1
   RUNG wire#powerrail
      { S7_Templates := "SrcType := String" } EQ_Contact(in1 := "Expected/Value_All".V, in2 := #Expected18)
   END_RUNG wire#w1
   RUNG wire#powerrail
      { S7_Templates := "SrcType := String" } EQ_Contact(in1 := "Expected/Value_All".V, in2 := #Expected19)
   END_RUNG wire#w1
   RUNG wire#powerrail
      { S7_Templates := "SrcType := String" } EQ_Contact(in1 := "Expected/Value_All".V, in2 := #Expected20)
   END_RUNG wire#w1
   // the same network as SCL:
   #On_Motor := ("Expected/Value_All".V = #Expected1) OR ("Expected/Value_All".V = #Expected2) OR ("Expected/Value_All".V = #Expected3) OR ("Expected/Value_All".V = #Expected4) OR ("Expected/Value_All".V = #Expected5) OR ("Expected/Value_All".V = #Expected6) OR ("Expected/Value_All".V = #Expected7) OR ("Expected/Value_All".V = #Expected8) OR ("Expected/Value_All".V = #Expected9) OR ("Expected/Value_All".V = #Expected10) OR ("Expected/Value_All".V = #Expected11) OR ("Expected/Value_All".V = #Expected12) OR ("Expected/Value_All".V = #Expected13) OR ("Expected/Value_All".V = #Expected14) OR ("Expected/Value_All".V = #Expected15) OR ("Expected/Value_All".V = #Expected16) OR ("Expected/Value_All".V = #Expected17) OR ("Expected/Value_All".V = #Expected18) OR ("Expected/Value_All".V = #Expected19) OR ("Expected/Value_All".V = #Expected20);
END_REGION
END_FUNCTION

// folder: System_In(จัดเก็บ)/Gripper System_In

FUNCTION_BLOCK "Gripper"   // FB2, LAD
{ S7_Optimized_Access := 'TRUE' }
VERSION : 0.1
   VAR_TEMP   // added for the SCL form of the ladder/FBD networks
      _w1 : Bool;
   END_VAR
BEGIN

REGION Network 1
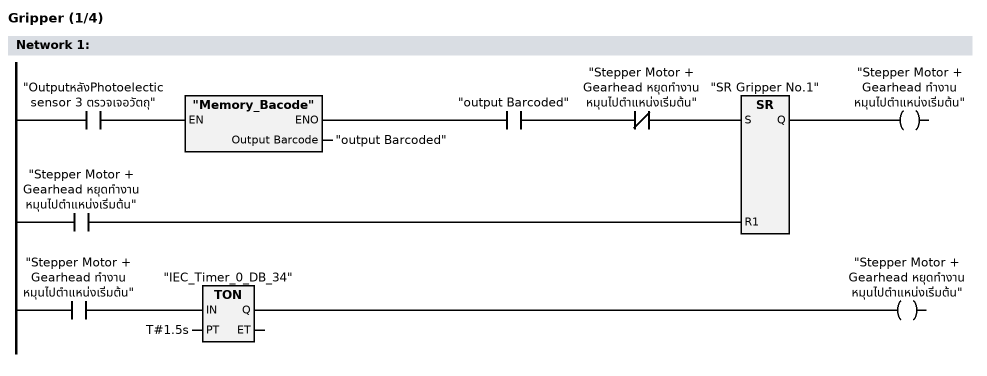
   "Memory_Bacode"(EN := "OutputหลังPhotoelectic sensor 3 ตรวจเจอวัตถุ",
                   "Output Barcode" => "output Barcoded",
                   ENO => #_w1);
   IF #_w1 AND "output Barcoded" AND NOT "Stepper Motor + Gearhead หยุดทำงาน หมุนไปตำแหน่งเริ่มต้น" THEN
       "SR Gripper No.1" := TRUE;   // SR flip-flop
   END_IF;
   IF "Stepper Motor + Gearhead หยุดทำงาน หมุนไปตำแหน่งเริ่มต้น" THEN "SR Gripper No.1" := FALSE; END_IF;
   "Stepper Motor + Gearhead ทำงาน หมุนไปตำแหน่งเริ่มต้น" := "SR Gripper No.1";
   "IEC_Timer_0_DB_34".TON(IN := "Stepper Motor + Gearhead ทำงาน หมุนไปตำแหน่งเริ่มต้น", PT := T#1.5s);
   "Stepper Motor + Gearhead หยุดทำงาน หมุนไปตำแหน่งเริ่มต้น" := "IEC_Timer_0_DB_34".Q;
END_REGION

REGION Network 2
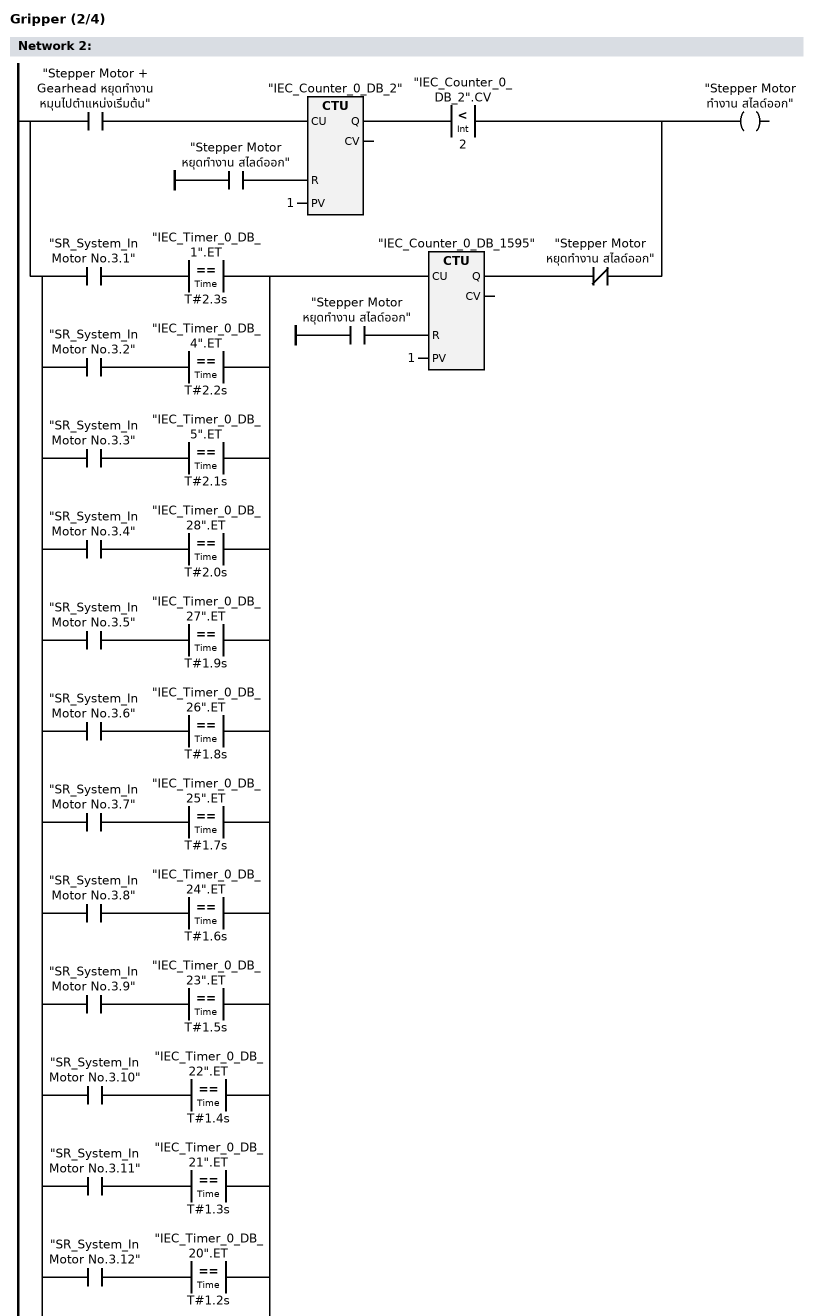
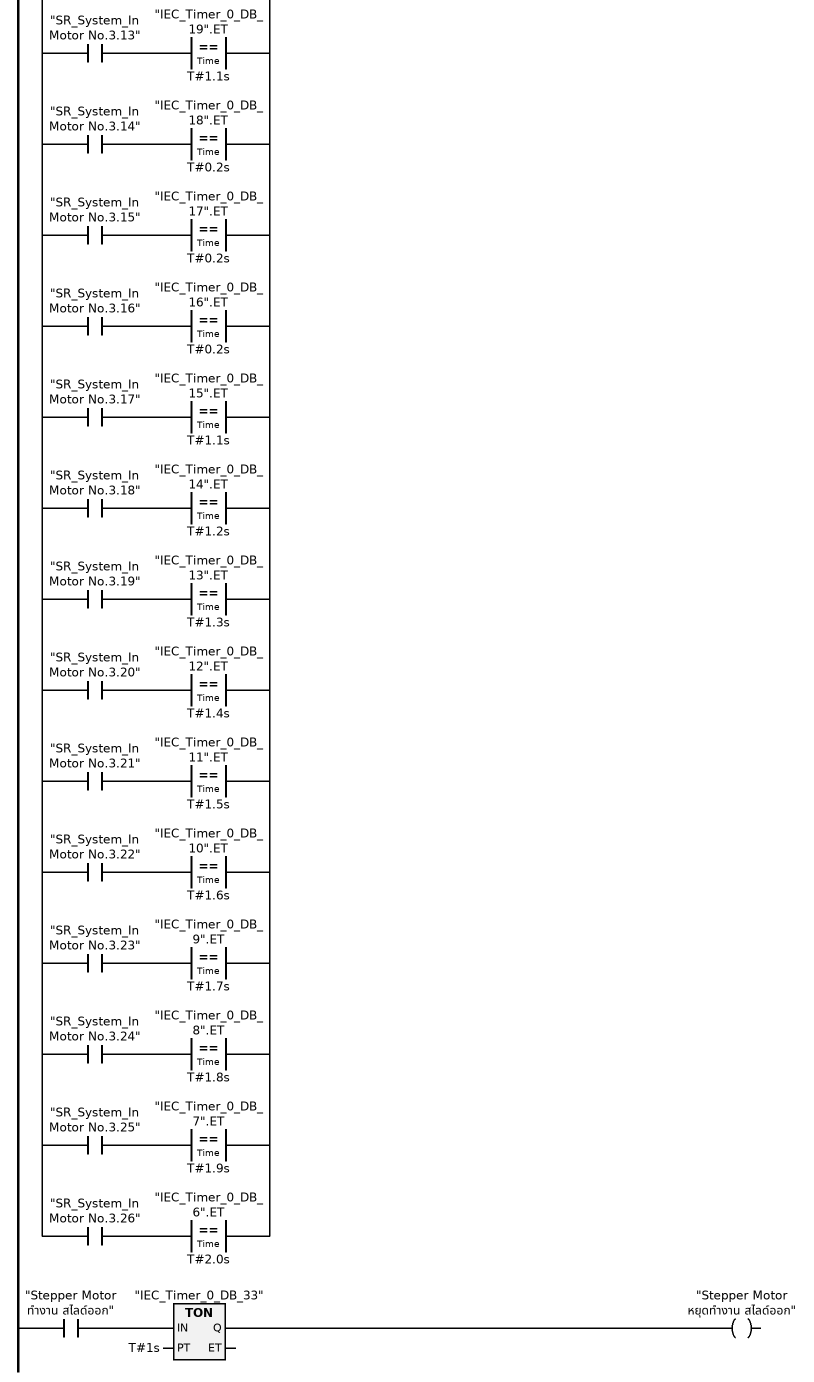
   "IEC_Counter_0_DB_2".CTU(CU := "Stepper Motor + Gearhead หยุดทำงาน หมุนไปตำแหน่งเริ่มต้น",
                           R := "Stepper Motor หยุดทำงาน สไลด์ออก",
                           PV := 1);
   "IEC_Counter_0_DB_1595".CTU(CU := ("SR_System_In Motor No.3.1" AND ("IEC_Timer_0_DB_1".ET = T#2.3s)) OR ("SR_System_In Motor No.3.2" AND ("IEC_Timer_0_DB_4".ET = T#2.2s)) OR ("SR_System_In Motor No.3.3" AND ("IEC_Timer_0_DB_5".ET = T#2.1s)) OR ("SR_System_In Motor No.3.4" AND ("IEC_Timer_0_DB_28".ET = T#2.0s)) OR ("SR_System_In Motor No.3.5" AND ("IEC_Timer_0_DB_27".ET = T#1.9s)) OR ("SR_System_In Motor No.3.6" AND ("IEC_Timer_0_DB_26".ET = T#1.8s)) OR ("SR_System_In Motor No.3.7" AND ("IEC_Timer_0_DB_25".ET = T#1.7s)) OR ("SR_System_In Motor No.3.8" AND ("IEC_Timer_0_DB_24".ET = T#1.6s)) OR ("SR_System_In Motor No.3.9" AND ("IEC_Timer_0_DB_23".ET = T#1.5s)) OR ("SR_System_In Motor No.3.10" AND ("IEC_Timer_0_DB_22".ET = T#1.4s)) OR ("SR_System_In Motor No.3.11" AND ("IEC_Timer_0_DB_21".ET = T#1.3s)) OR ("SR_System_In Motor No.3.12" AND ("IEC_Timer_0_DB_20".ET = T#1.2s)) OR ("SR_System_In Motor No.3.13" AND ("IEC_Timer_0_DB_19".ET = T#1.1s)) OR ("SR_System_In Motor No.3.14" AND ("IEC_Timer_0_DB_18".ET = T#0.2s)) OR ("SR_System_In Motor No.3.15" AND ("IEC_Timer_0_DB_17".ET = T#0.2s)) OR ("SR_System_In Motor No.3.16" AND ("IEC_Timer_0_DB_16".ET = T#0.2s)) OR ("SR_System_In Motor No.3.17" AND ("IEC_Timer_0_DB_15".ET = T#1.1s)) OR ("SR_System_In Motor No.3.18" AND ("IEC_Timer_0_DB_14".ET = T#1.2s)) OR ("SR_System_In Motor No.3.19" AND ("IEC_Timer_0_DB_13".ET = T#1.3s)) OR ("SR_System_In Motor No.3.20" AND ("IEC_Timer_0_DB_12".ET = T#1.4s)) OR ("SR_System_In Motor No.3.21" AND ("IEC_Timer_0_DB_11".ET = T#1.5s)) OR ("SR_System_In Motor No.3.22" AND ("IEC_Timer_0_DB_10".ET = T#1.6s)) OR ("SR_System_In Motor No.3.23" AND ("IEC_Timer_0_DB_9".ET = T#1.7s)) OR ("SR_System_In Motor No.3.24" AND ("IEC_Timer_0_DB_8".ET = T#1.8s)) OR ("SR_System_In Motor No.3.25" AND ("IEC_Timer_0_DB_7".ET = T#1.9s)) OR ("SR_System_In Motor No.3.26" AND ("IEC_Timer_0_DB_6".ET = T#2.0s)),
                           R := "Stepper Motor หยุดทำงาน สไลด์ออก",
                           PV := 1);
   "Stepper Motor ทำงาน สไลด์ออก" := ("IEC_Counter_0_DB_2".Q AND ("IEC_Counter_0_DB_2".CV < 2)) OR ("IEC_Counter_0_DB_1595".Q AND NOT "Stepper Motor หยุดทำงาน สไลด์ออก");
   "IEC_Timer_0_DB_33".TON(IN := "Stepper Motor ทำงาน สไลด์ออก", PT := T#1s);
   "Stepper Motor หยุดทำงาน สไลด์ออก" := "IEC_Timer_0_DB_33".Q;
END_REGION

REGION Network 3
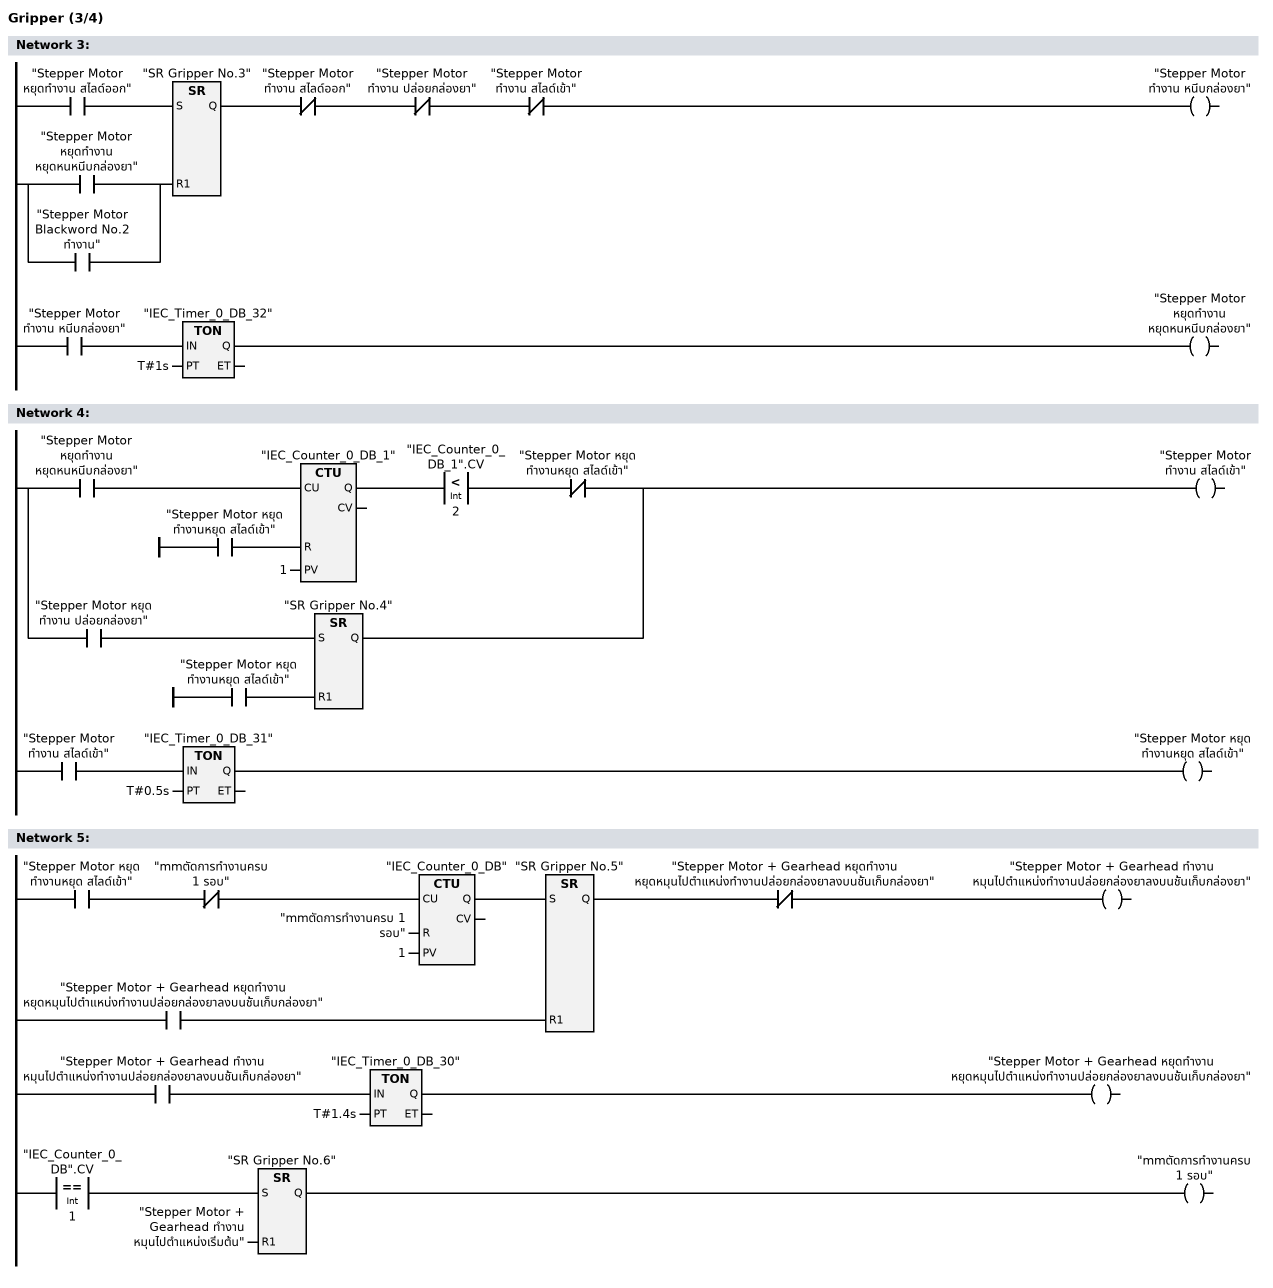
   IF "Stepper Motor หยุดทำงาน สไลด์ออก" THEN
       "SR Gripper No.3" := TRUE;   // SR flip-flop
   END_IF;
   IF "Stepper Motor หยุดทำงาน หยุดหนหนีบกล่องยา" OR "Stepper Motor Blackword No.2 ทำงาน" THEN
       "SR Gripper No.3" := FALSE;
   END_IF;
   "Stepper Motor ทำงาน หนีบกล่องยา" := "SR Gripper No.3" AND NOT "Stepper Motor ทำงาน สไลด์ออก" AND NOT "Stepper Motor ทำงาน ปล่อยกล่องยา" AND NOT "Stepper Motor ทำงาน สไลด์เข้า";
   "IEC_Timer_0_DB_32".TON(IN := "Stepper Motor ทำงาน หนีบกล่องยา", PT := T#1s);
   "Stepper Motor หยุดทำงาน หยุดหนหนีบกล่องยา" := "IEC_Timer_0_DB_32".Q;
END_REGION

REGION Network 4
   "IEC_Counter_0_DB_1".CTU(CU := "Stepper Motor หยุดทำงาน หยุดหนหนีบกล่องยา",
                           R := "Stepper Motor หยุด ทำงานหยุด สไลด์เข้า",
                           PV := 1);
   IF "Stepper Motor หยุด ทำงาน ปล่อยกล่องยา" THEN
       "SR Gripper No.4" := TRUE;   // SR flip-flop
   END_IF;
   IF "Stepper Motor หยุด ทำงานหยุด สไลด์เข้า" THEN "SR Gripper No.4" := FALSE; END_IF;
   "Stepper Motor ทำงาน สไลด์เข้า" := ("IEC_Counter_0_DB_1".Q AND ("IEC_Counter_0_DB_1".CV < 2) AND NOT "Stepper Motor หยุด ทำงานหยุด สไลด์เข้า") OR "SR Gripper No.4";
   "IEC_Timer_0_DB_31".TON(IN := "Stepper Motor ทำงาน สไลด์เข้า", PT := T#0.5s);
   "Stepper Motor หยุด ทำงานหยุด สไลด์เข้า" := "IEC_Timer_0_DB_31".Q;
END_REGION

REGION Network 5
   "IEC_Counter_0_DB".CTU(CU := "Stepper Motor หยุด ทำงานหยุด สไลด์เข้า" AND NOT "mmตัดการทำงานครบ 1 รอบ",
                          R := "mmตัดการทำงานครบ 1 รอบ",
                          PV := 1);
   IF "IEC_Counter_0_DB".Q THEN
       "SR Gripper No.5" := TRUE;   // SR flip-flop
   END_IF;
   IF "Stepper Motor + Gearhead หยุดทำงาน หยุดหมุนไปตำแหน่งทำงานปล่อยกล่องยาลงบนชั้นเก็บกล่องยา" THEN
       "SR Gripper No.5" := FALSE;
   END_IF;
   "Stepper Motor + Gearhead ทำงาน หมุนไปตำแหน่งทำงานปล่อยกล่องยาลงบนชั้นเก็บกล่องยา" := "SR Gripper No.5" AND NOT "Stepper Motor + Gearhead หยุดทำงาน หยุดหมุนไปตำแหน่งทำงานปล่อยกล่องยาลงบนชั้นเก็บกล่องยา";
   "IEC_Timer_0_DB_30".TON(IN := "Stepper Motor + Gearhead ทำงาน หมุนไปตำแหน่งทำงานปล่อยกล่องยาลงบนชั้นเก็บกล่องยา",
                           PT := T#1.4s);
   "Stepper Motor + Gearhead หยุดทำงาน หยุดหมุนไปตำแหน่งทำงานปล่อยกล่องยาลงบนชั้นเก็บกล่องยา" := "IEC_Timer_0_DB_30".Q;
   IF "IEC_Counter_0_DB".CV = 1 THEN
       "SR Gripper No.6" := TRUE;   // SR flip-flop
   END_IF;
   IF "Stepper Motor + Gearhead ทำงาน หมุนไปตำแหน่งเริ่มต้น" THEN "SR Gripper No.6" := FALSE; END_IF;
   "mmตัดการทำงานครบ 1 รอบ" := "SR Gripper No.6";
END_REGION

REGION Network 6
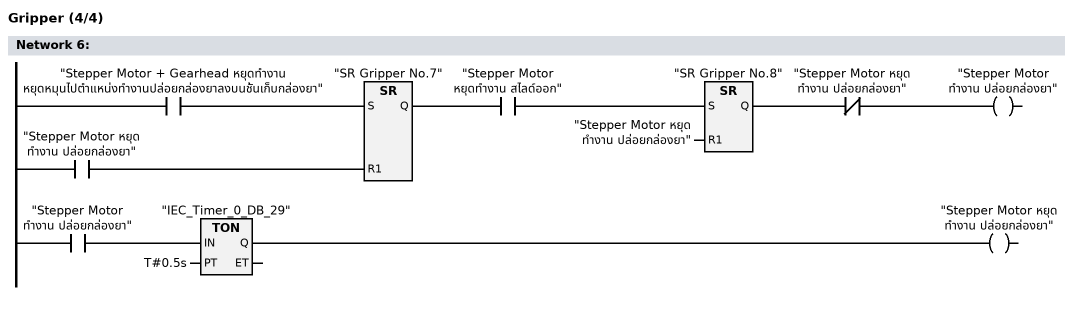
   IF "Stepper Motor + Gearhead หยุดทำงาน หยุดหมุนไปตำแหน่งทำงานปล่อยกล่องยาลงบนชั้นเก็บกล่องยา" THEN
       "SR Gripper No.7" := TRUE;   // SR flip-flop
   END_IF;
   IF "Stepper Motor หยุด ทำงาน ปล่อยกล่องยา" THEN "SR Gripper No.7" := FALSE; END_IF;
   IF "SR Gripper No.7" AND "Stepper Motor หยุดทำงาน สไลด์ออก" THEN
       "SR Gripper No.8" := TRUE;   // SR flip-flop
   END_IF;
   IF "Stepper Motor หยุด ทำงาน ปล่อยกล่องยา" THEN "SR Gripper No.8" := FALSE; END_IF;
   "Stepper Motor ทำงาน ปล่อยกล่องยา" := "SR Gripper No.8" AND NOT "Stepper Motor หยุด ทำงาน ปล่อยกล่องยา";
   "IEC_Timer_0_DB_29".TON(IN := "Stepper Motor ทำงาน ปล่อยกล่องยา", PT := T#0.5s);
   "Stepper Motor หยุด ทำงาน ปล่อยกล่องยา" := "IEC_Timer_0_DB_29".Q;
END_REGION
END_FUNCTION_BLOCK

FUNCTION "Motor ถึงตำแหน่งเป้าหมาย" : Void   // FC6, LAD
{ S7_Optimized_Access := 'TRUE' }
VERSION : 0.1
   VAR_OUTPUT
      Output : Bool;
   END_VAR
BEGIN

REGION Network 1
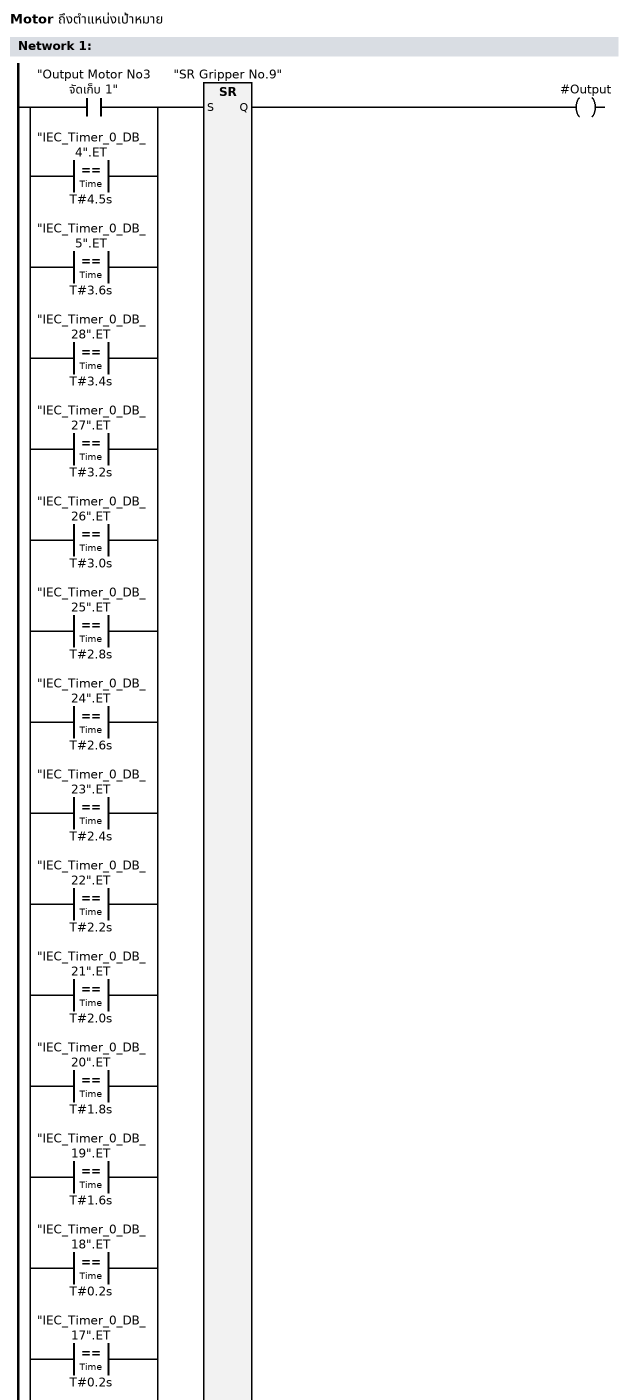
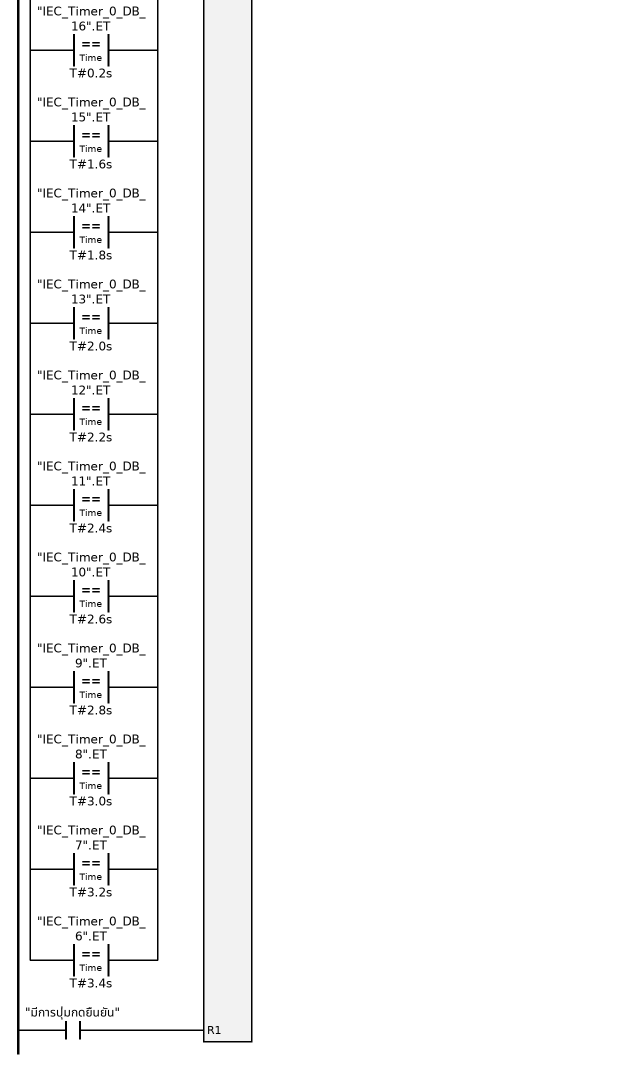
   RUNG wire#powerrail
      Contact( "Output Motor No3 จัดเก็บ 1" )
      wire#w1
      S_SR(operand := "SR Gripper No.9", r1 := wire#w2)
      Coil( #Output )
   END_RUNG
   RUNG wire#powerrail
      { S7_Templates := "SrcType := Time" } EQ_Contact(in1 := "IEC_Timer_0_DB_4".ET, in2 := T#4.5s)
   END_RUNG wire#w1
   RUNG wire#powerrail
      { S7_Templates := "SrcType := Time" } EQ_Contact(in1 := "IEC_Timer_0_DB_5".ET, in2 := T#3.6s)
   END_RUNG wire#w1
   RUNG wire#powerrail
      { S7_Templates := "SrcType := Time" } EQ_Contact(in1 := "IEC_Timer_0_DB_28".ET, in2 := T#3.4s)
   END_RUNG wire#w1
   RUNG wire#powerrail
      { S7_Templates := "SrcType := Time" } EQ_Contact(in1 := "IEC_Timer_0_DB_27".ET, in2 := T#3.2s)
   END_RUNG wire#w1
   RUNG wire#powerrail
      { S7_Templates := "SrcType := Time" } EQ_Contact(in1 := "IEC_Timer_0_DB_26".ET, in2 := T#3.0s)
   END_RUNG wire#w1
   RUNG wire#powerrail
      { S7_Templates := "SrcType := Time" } EQ_Contact(in1 := "IEC_Timer_0_DB_25".ET, in2 := T#2.8s)
   END_RUNG wire#w1
   RUNG wire#powerrail
      { S7_Templates := "SrcType := Time" } EQ_Contact(in1 := "IEC_Timer_0_DB_24".ET, in2 := T#2.6s)
   END_RUNG wire#w1
   RUNG wire#powerrail
      { S7_Templates := "SrcType := Time" } EQ_Contact(in1 := "IEC_Timer_0_DB_23".ET, in2 := T#2.4s)
   END_RUNG wire#w1
   RUNG wire#powerrail
      { S7_Templates := "SrcType := Time" } EQ_Contact(in1 := "IEC_Timer_0_DB_22".ET, in2 := T#2.2s)
   END_RUNG wire#w1
   RUNG wire#powerrail
      { S7_Templates := "SrcType := Time" } EQ_Contact(in1 := "IEC_Timer_0_DB_21".ET, in2 := T#2.0s)
   END_RUNG wire#w1
   RUNG wire#powerrail
      { S7_Templates := "SrcType := Time" } EQ_Contact(in1 := "IEC_Timer_0_DB_20".ET, in2 := T#1.8s)
   END_RUNG wire#w1
   RUNG wire#powerrail
      { S7_Templates := "SrcType := Time" } EQ_Contact(in1 := "IEC_Timer_0_DB_19".ET, in2 := T#1.6s)
   END_RUNG wire#w1
   RUNG wire#powerrail
      { S7_Templates := "SrcType := Time" } EQ_Contact(in1 := "IEC_Timer_0_DB_18".ET, in2 := T#0.2s)
   END_RUNG wire#w1
   RUNG wire#powerrail
      { S7_Templates := "SrcType := Time" } EQ_Contact(in1 := "IEC_Timer_0_DB_17".ET, in2 := T#0.2s)
   END_RUNG wire#w1
   RUNG wire#powerrail
      { S7_Templates := "SrcType := Time" } EQ_Contact(in1 := "IEC_Timer_0_DB_16".ET, in2 := T#0.2s)
   END_RUNG wire#w1
   RUNG wire#powerrail
      { S7_Templates := "SrcType := Time" } EQ_Contact(in1 := "IEC_Timer_0_DB_15".ET, in2 := T#1.6s)
   END_RUNG wire#w1
   RUNG wire#powerrail
      { S7_Templates := "SrcType := Time" } EQ_Contact(in1 := "IEC_Timer_0_DB_14".ET, in2 := T#1.8s)
   END_RUNG wire#w1
   RUNG wire#powerrail
      { S7_Templates := "SrcType := Time" } EQ_Contact(in1 := "IEC_Timer_0_DB_13".ET, in2 := T#2.0s)
   END_RUNG wire#w1
   RUNG wire#powerrail
      { S7_Templates := "SrcType := Time" } EQ_Contact(in1 := "IEC_Timer_0_DB_12".ET, in2 := T#2.2s)
   END_RUNG wire#w1
   RUNG wire#powerrail
      { S7_Templates := "SrcType := Time" } EQ_Contact(in1 := "IEC_Timer_0_DB_11".ET, in2 := T#2.4s)
   END_RUNG wire#w1
   RUNG wire#powerrail
      { S7_Templates := "SrcType := Time" } EQ_Contact(in1 := "IEC_Timer_0_DB_10".ET, in2 := T#2.6s)
   END_RUNG wire#w1
   RUNG wire#powerrail
      { S7_Templates := "SrcType := Time" } EQ_Contact(in1 := "IEC_Timer_0_DB_9".ET, in2 := T#2.8s)
   END_RUNG wire#w1
   RUNG wire#powerrail
      { S7_Templates := "SrcType := Time" } EQ_Contact(in1 := "IEC_Timer_0_DB_8".ET, in2 := T#3.0s)
   END_RUNG wire#w1
   RUNG wire#powerrail
      { S7_Templates := "SrcType := Time" } EQ_Contact(in1 := "IEC_Timer_0_DB_7".ET, in2 := T#3.2s)
   END_RUNG wire#w1
   RUNG wire#powerrail
      { S7_Templates := "SrcType := Time" } EQ_Contact(in1 := "IEC_Timer_0_DB_6".ET, in2 := T#3.4s)
   END_RUNG wire#w1
   RUNG wire#powerrail
      Contact( "มีการปุ่มกดยืนยัน" )
   END_RUNG wire#w2
   // the same network as SCL:
   IF "Output Motor No3 จัดเก็บ 1" OR ("IEC_Timer_0_DB_4".ET = T#4.5s) OR ("IEC_Timer_0_DB_5".ET = T#3.6s) OR ("IEC_Timer_0_DB_28".ET = T#3.4s) OR ("IEC_Timer_0_DB_27".ET = T#3.2s) OR ("IEC_Timer_0_DB_26".ET = T#3.0s) OR ("IEC_Timer_0_DB_25".ET = T#2.8s) OR ("IEC_Timer_0_DB_24".ET = T#2.6s) OR ("IEC_Timer_0_DB_23".ET = T#2.4s) OR ("IEC_Timer_0_DB_22".ET = T#2.2s) OR ("IEC_Timer_0_DB_21".ET = T#2.0s) OR ("IEC_Timer_0_DB_20".ET = T#1.8s) OR ("IEC_Timer_0_DB_19".ET = T#1.6s) OR ("IEC_Timer_0_DB_18".ET = T#0.2s) OR ("IEC_Timer_0_DB_17".ET = T#0.2s) OR ("IEC_Timer_0_DB_16".ET = T#0.2s) OR ("IEC_Timer_0_DB_15".ET = T#1.6s) OR ("IEC_Timer_0_DB_14".ET = T#1.8s) OR ("IEC_Timer_0_DB_13".ET = T#2.0s) OR ("IEC_Timer_0_DB_12".ET = T#2.2s) OR ("IEC_Timer_0_DB_11".ET = T#2.4s) OR ("IEC_Timer_0_DB_10".ET = T#2.6s) OR ("IEC_Timer_0_DB_9".ET = T#2.8s) OR ("IEC_Timer_0_DB_8".ET = T#3.0s) OR ("IEC_Timer_0_DB_7".ET = T#3.2s) OR ("IEC_Timer_0_DB_6".ET = T#3.4s) THEN
       "SR Gripper No.9" := TRUE;   // SR flip-flop
   END_IF;
   IF "มีการปุ่มกดยืนยัน" THEN "SR Gripper No.9" := FALSE; END_IF;
   #Output := "SR Gripper No.9";
END_REGION
END_FUNCTION

FUNCTION "test หลังเคลื่อนที่มาตำแหน่งปล่อยกล่องยา" : Void   // FC7, LAD
{ S7_Optimized_Access := 'TRUE' }
VERSION : 0.1
BEGIN

REGION Network 1
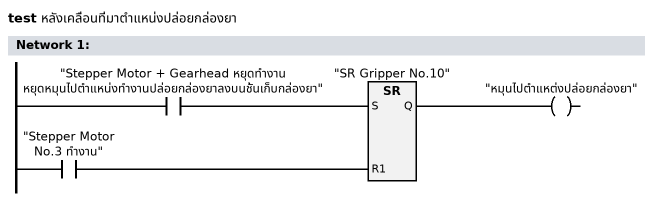
   RUNG wire#powerrail
      Contact( "Stepper Motor + Gearhead หยุดทำงาน หยุดหมุนไปตำแหน่งทำงานปล่อยกล่องยาลงบนชั้นเก็บกล่องยา" )
      S_SR(operand := "SR Gripper No.10", r1 := wire#w1)
      Coil( "หมุนไปตำแหต่งปล่อยกล่องยา" )
   END_RUNG
   RUNG wire#powerrail
      Contact( "Stepper Motor No.3 ทำงาน" )
   END_RUNG wire#w1
   // the same network as SCL:
   IF "Stepper Motor + Gearhead หยุดทำงาน หยุดหมุนไปตำแหน่งทำงานปล่อยกล่องยาลงบนชั้นเก็บกล่องยา" THEN
       "SR Gripper No.10" := TRUE;   // SR flip-flop
   END_IF;
   IF "Stepper Motor No.3 ทำงาน" THEN "SR Gripper No.10" := FALSE; END_IF;
   "หมุนไปตำแหต่งปล่อยกล่องยา" := "SR Gripper No.10";
END_REGION
END_FUNCTION

// folder: System_In(จัดเก็บ)/Step motor No.1,No.2

FUNCTION_BLOCK "Step motor ขึ่น-ลง ตามแกน y No.1,No.2_Forword"   // FB1, LAD
{ S7_Optimized_Access := 'TRUE' }
VERSION : 0.1
   VAR_INPUT
      Value : String;
      "TIME ที่ใช้ไป BOX.1-BOX.26" : Time;
      "TIME ที่ใช้ไป BOX.27-BOX.52" : Time;
      "TIME ที่ใช้ไป BOX.53-BOX.78" : Time;
      "TIME ที่ใช้ไป BOX.79-BOX.104" : Time;
      "TIME ที่ใช้ไป BOX.105-BOX.130" : Time;
      "TIME ที่ใช้ไป BOX.131-BOX.156" : Time;
      "TIME ที่ใช้ไป BOX.157-BOX.182" : Time;
      "TIME ที่ใช้ไป BOX.183-BOX.208" : Time;
      "TIME ที่ใช้ไป BOX.209-BOX.234" : Time;
      "TIME ที่ใช้ไป BOX.235-BOX.260" : Time;
      "TIME ที่ใช้ไป BOX.261-BOX.286" : Time;
      "TIME ที่ใช้ไป BOX.287-BOX.312" : Time;
      "TIME ที่ใช้ไป BOX.313-BOX.338" : Time;
      "TIME ที่ใช้ไป BOX.339-BOX.364" : Time;
      "TIME ที่ใช้ไป BOX.365-BOX.390" : Time;
      "TIME ที่ใช้ไป BOX.391-BOX.416" : Time;
      "TIME ที่ใช้ไป BOX.417-BOX.442" : Time;
      "TIME ที่ใช้ไป BOX.443-BOX.468" : Time;
      "TIME ที่ใช้ไป BOX.469-BOX.494" : Time;
      "TIME ที่ใช้ไป BOX.495-BOX.520" : Time;
   END_VAR
   VAR_IN_OUT
      "Stepper Motor  ทำงาน" : Bool;
   END_VAR
   VAR_TEMP   // added for the SCL form of the ladder/FBD networks
      _w1 : Bool;
      _w2 : Bool;
      _w3 : Bool;
      _w4 : Bool;
      _w5 : Bool;
      _w6 : Bool;
      _w7 : Bool;
      _w8 : Bool;
      _w9 : Bool;
      _w10 : Bool;
      _w11 : Bool;
      _w12 : Bool;
      _w13 : Bool;
      _w14 : Bool;
      _w15 : Bool;
      _w16 : Bool;
      _w17 : Bool;
      _w18 : Bool;
      _w19 : Bool;
      _w20 : Bool;
      _w21 : Bool;
      _w22 : Bool;
      _w23 : Bool;
      _w24 : Bool;
      _w25 : Bool;
      _w26 : Bool;
      _w27 : Bool;
      _w28 : Bool;
      _w29 : Bool;
      _w30 : Bool;
      _w31 : Bool;
      _w32 : Bool;
      _w33 : Bool;
      _w34 : Bool;
      _w35 : Bool;
      _w36 : Bool;
      _w37 : Bool;
      _w38 : Bool;
      _w39 : Bool;
      _w40 : Bool;
   END_VAR
BEGIN

REGION Network 1
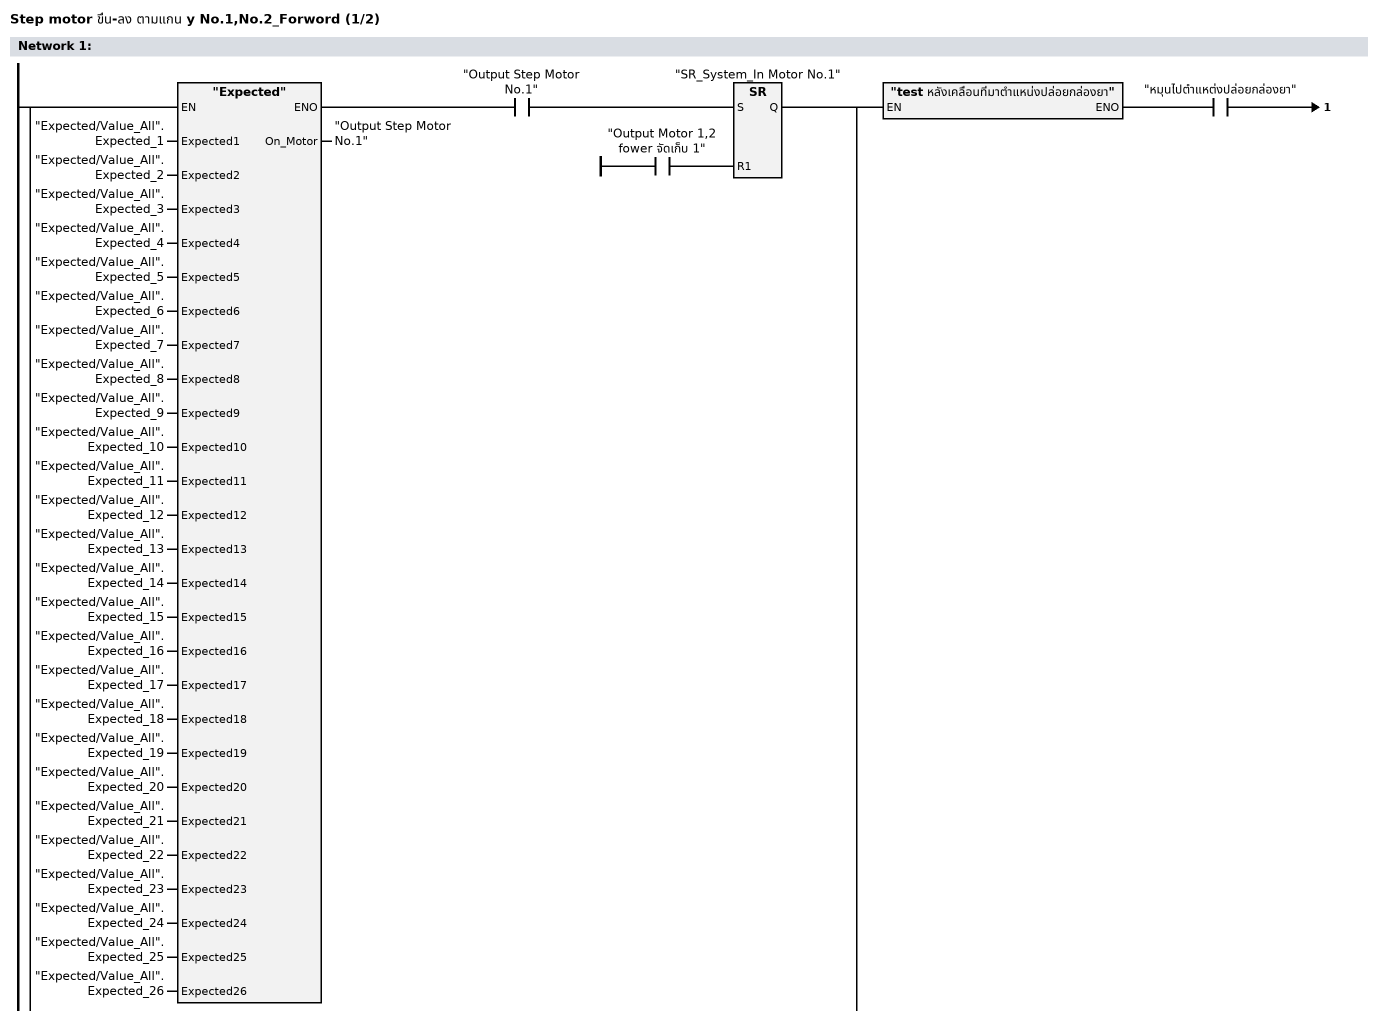
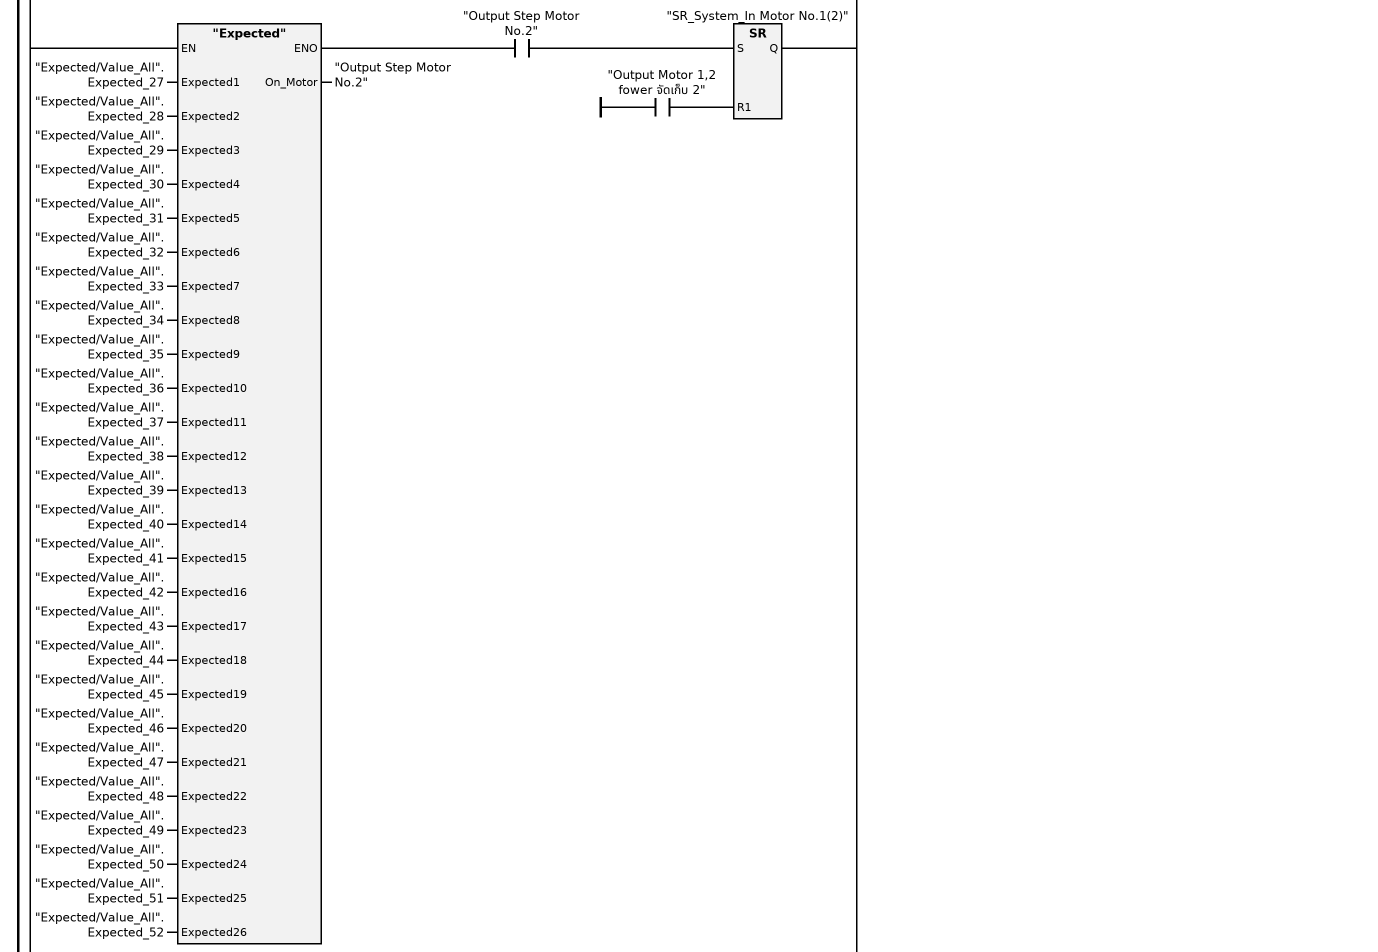
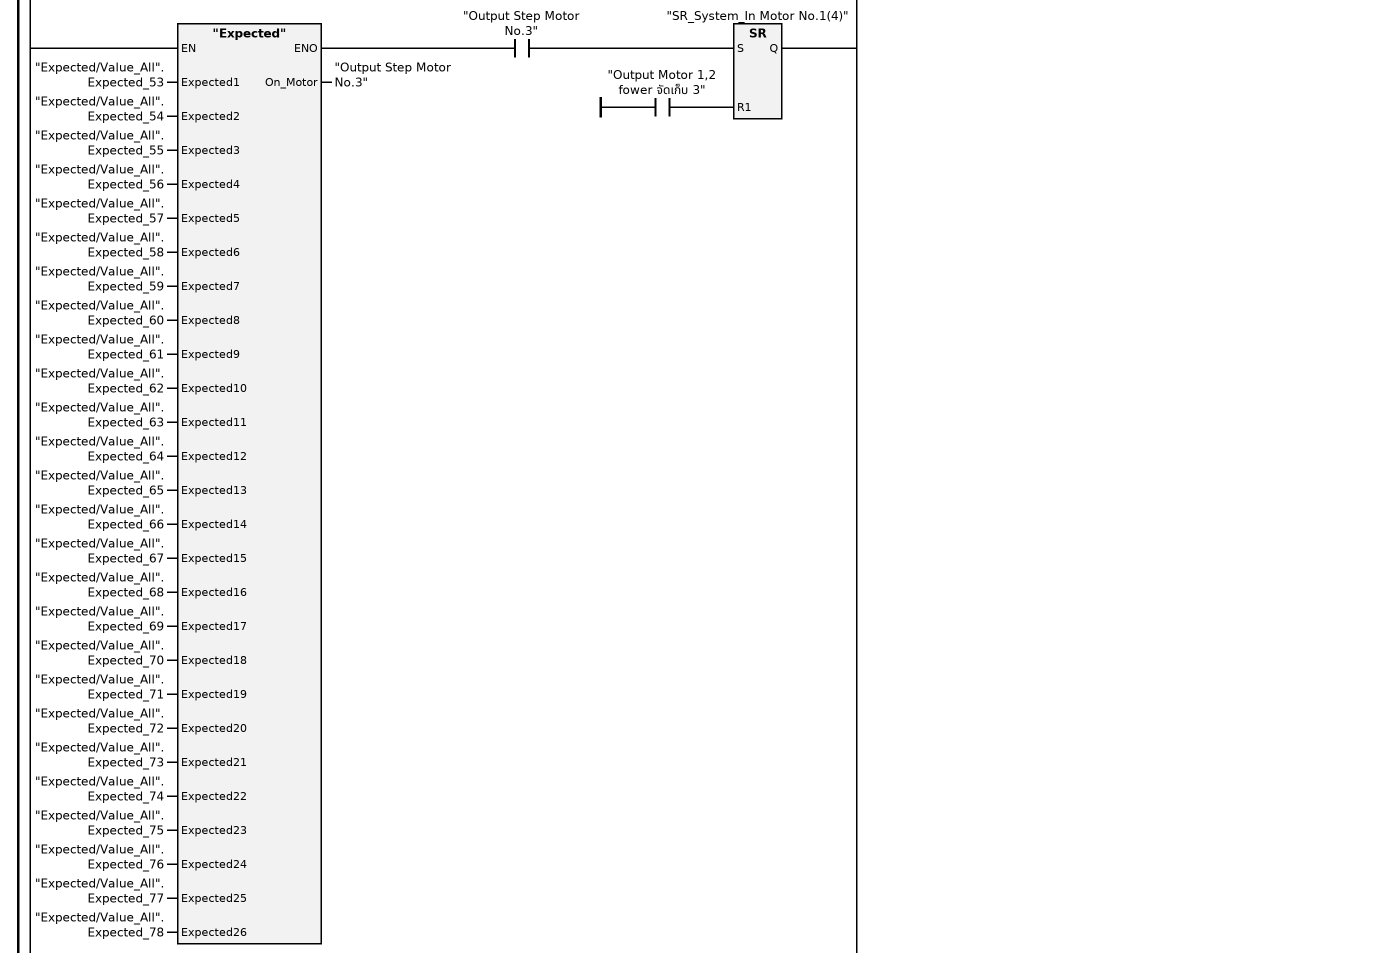
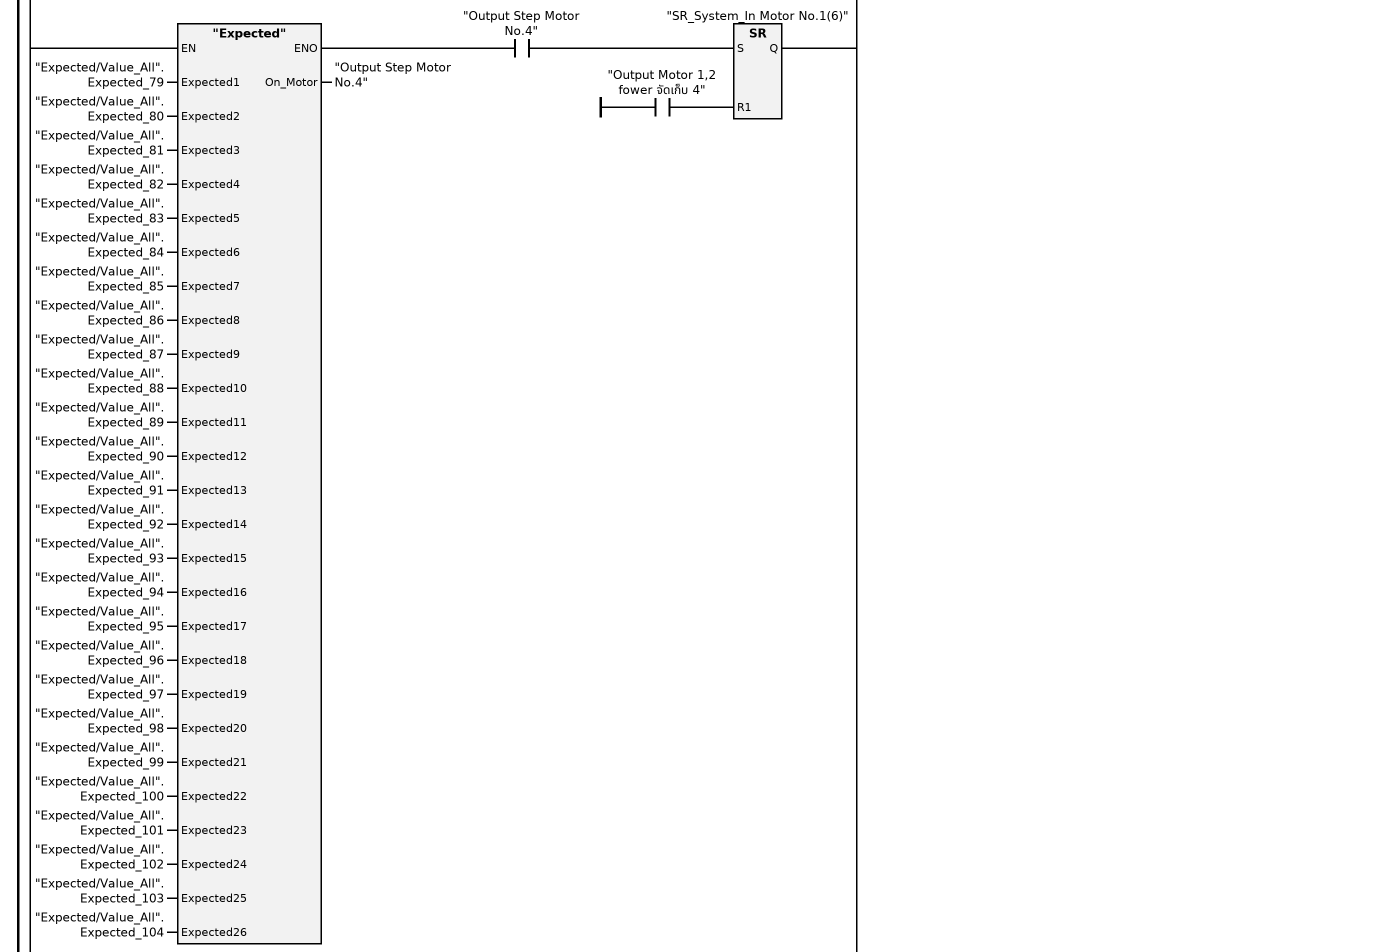
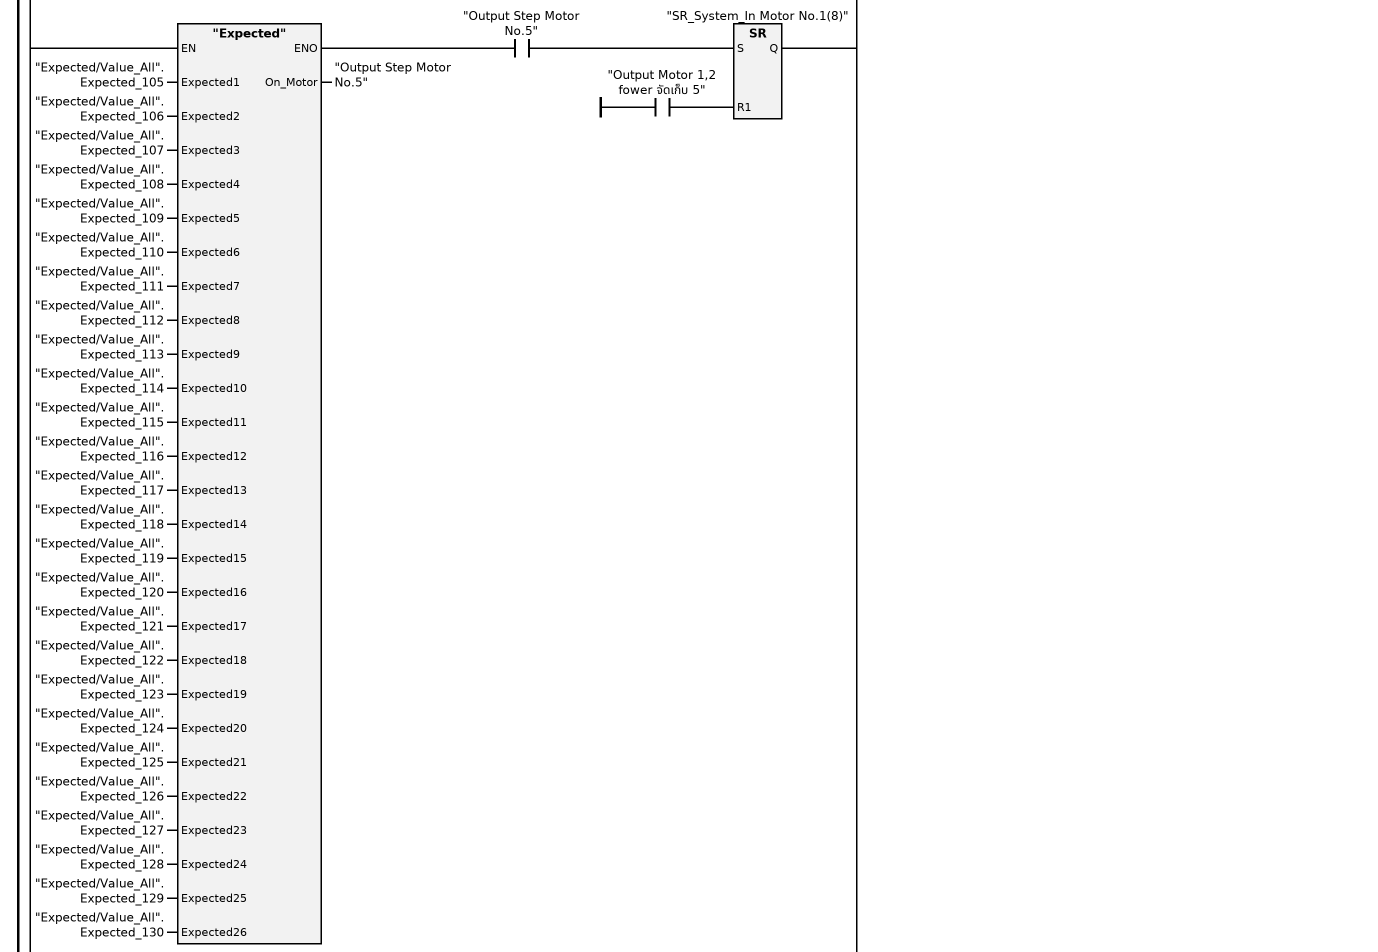
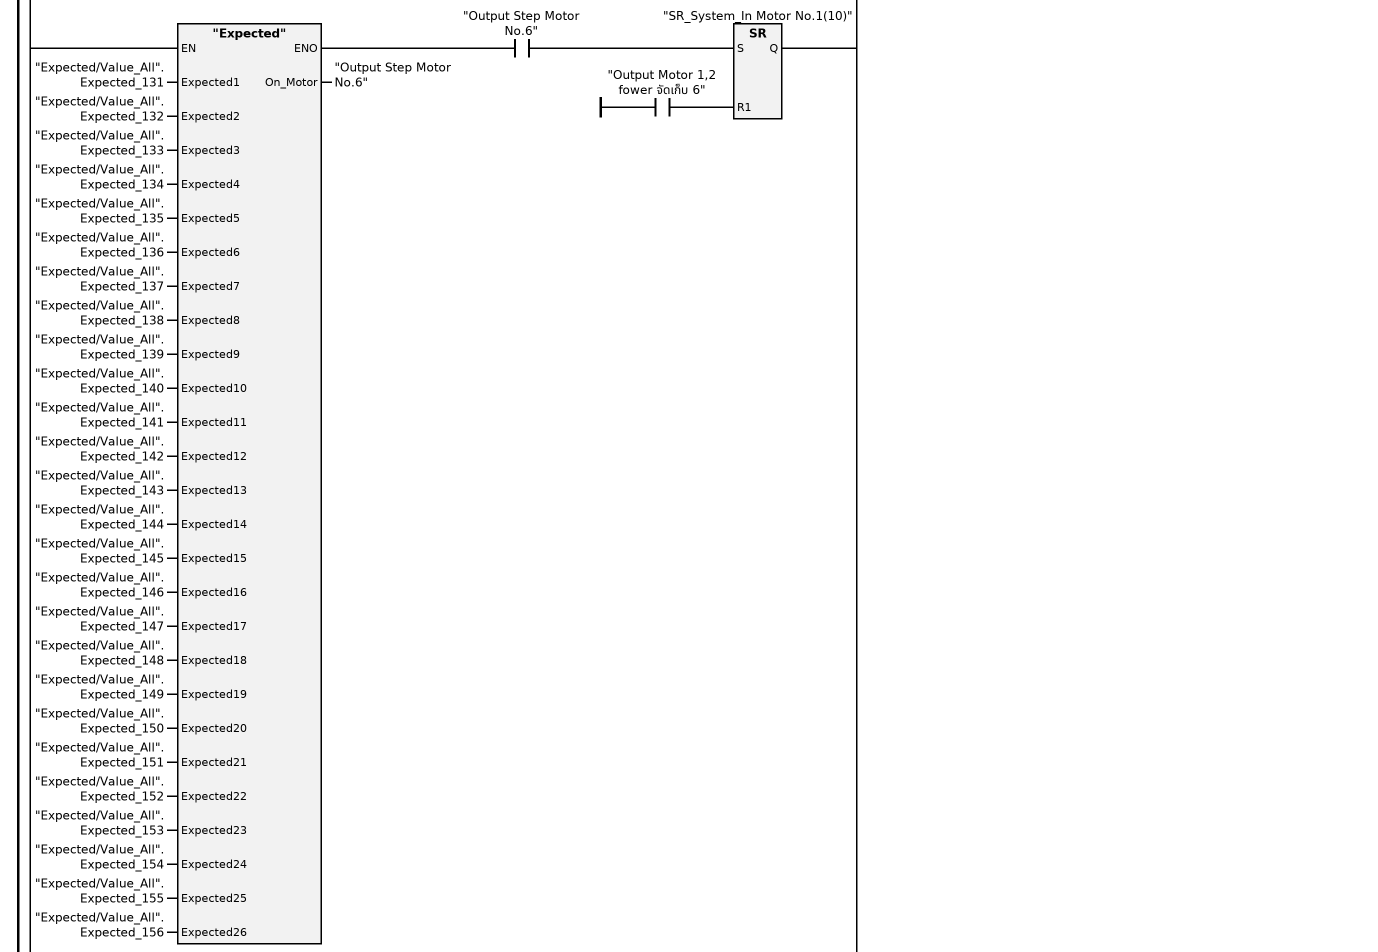
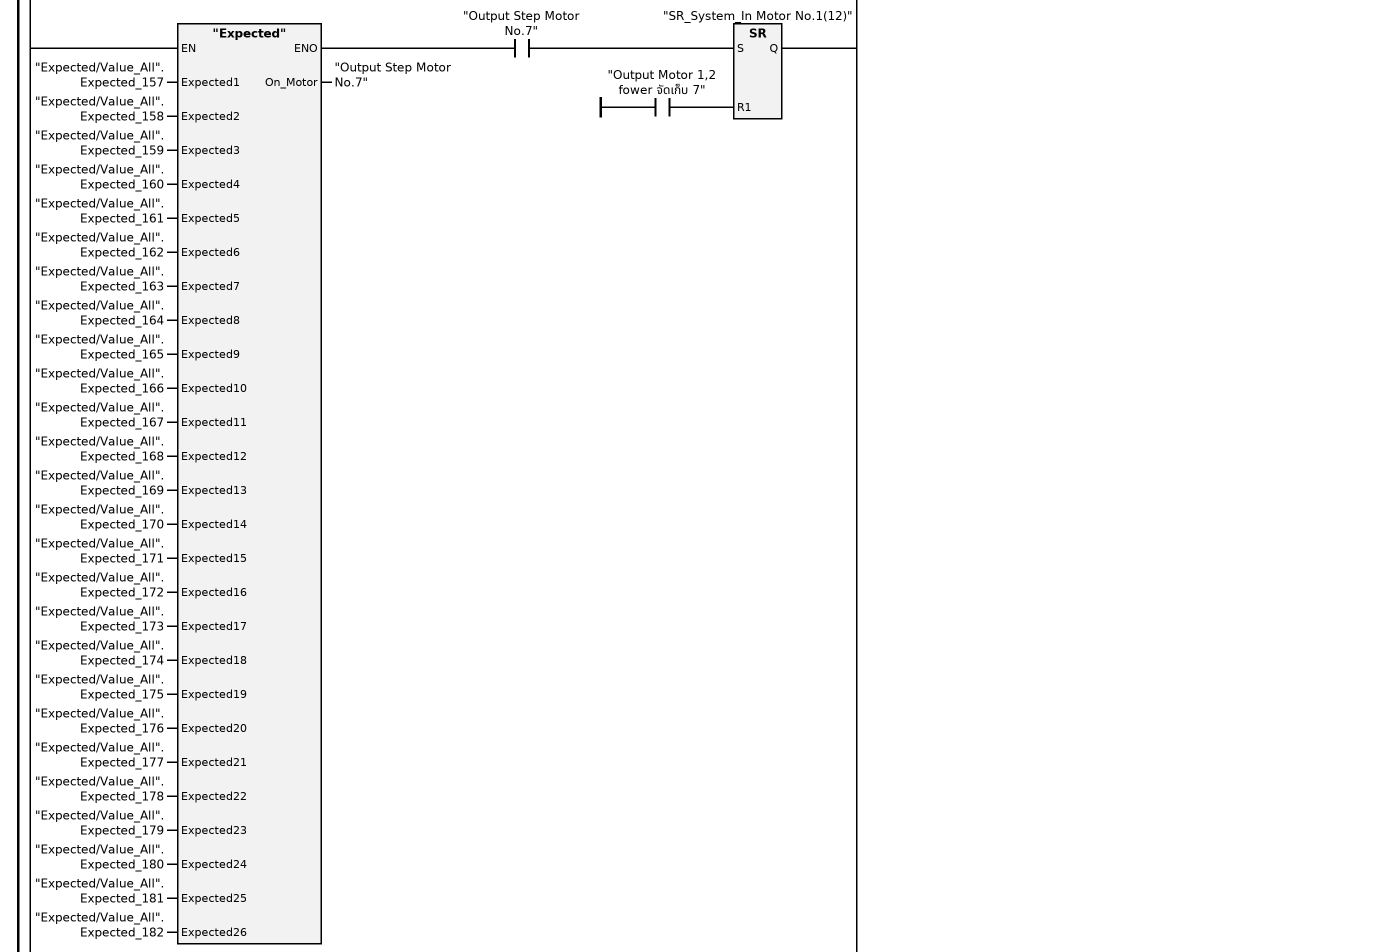
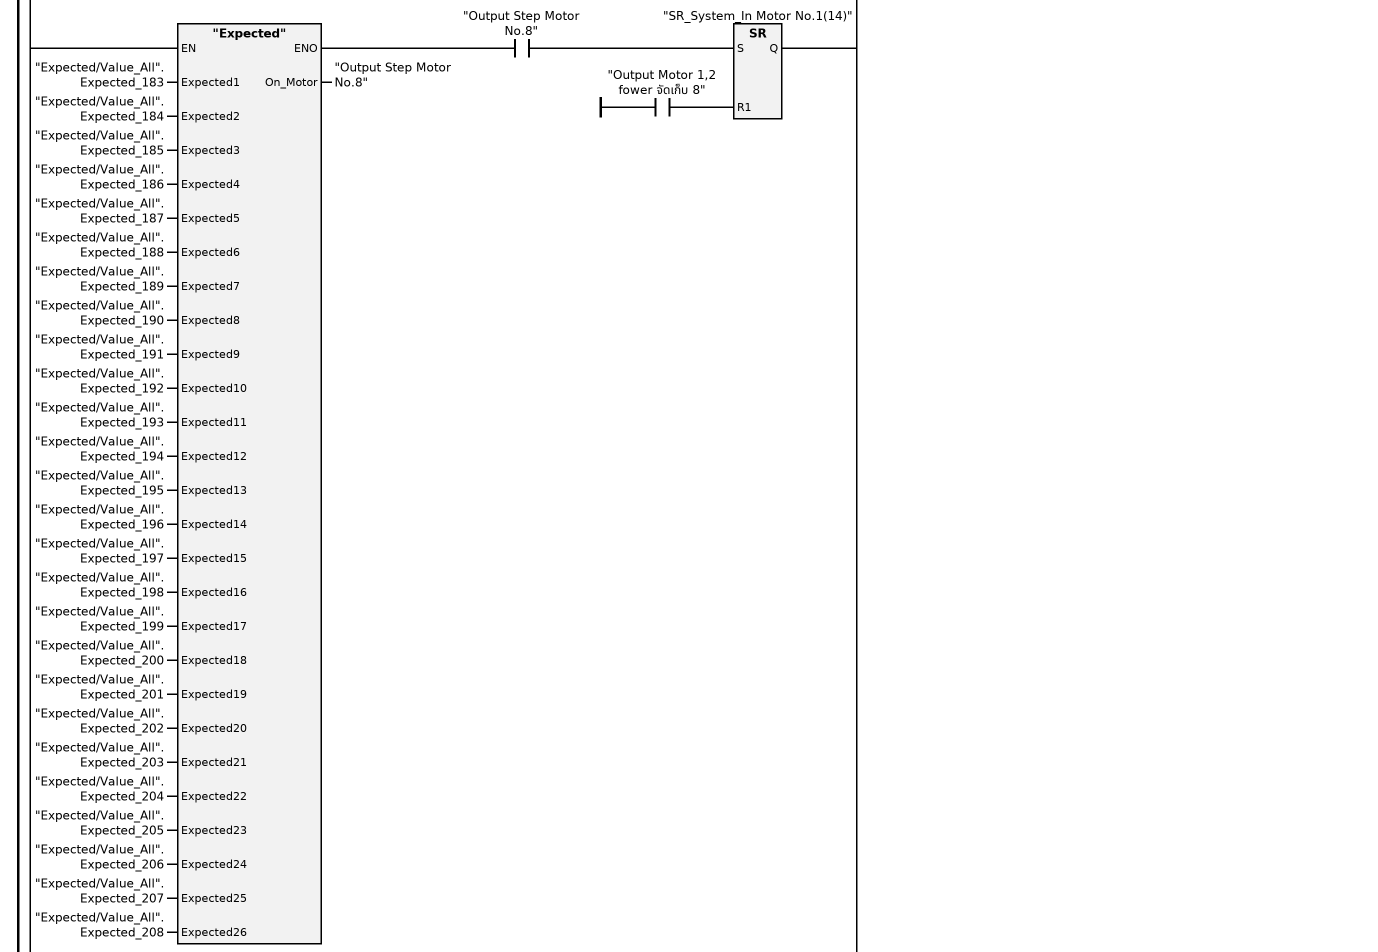
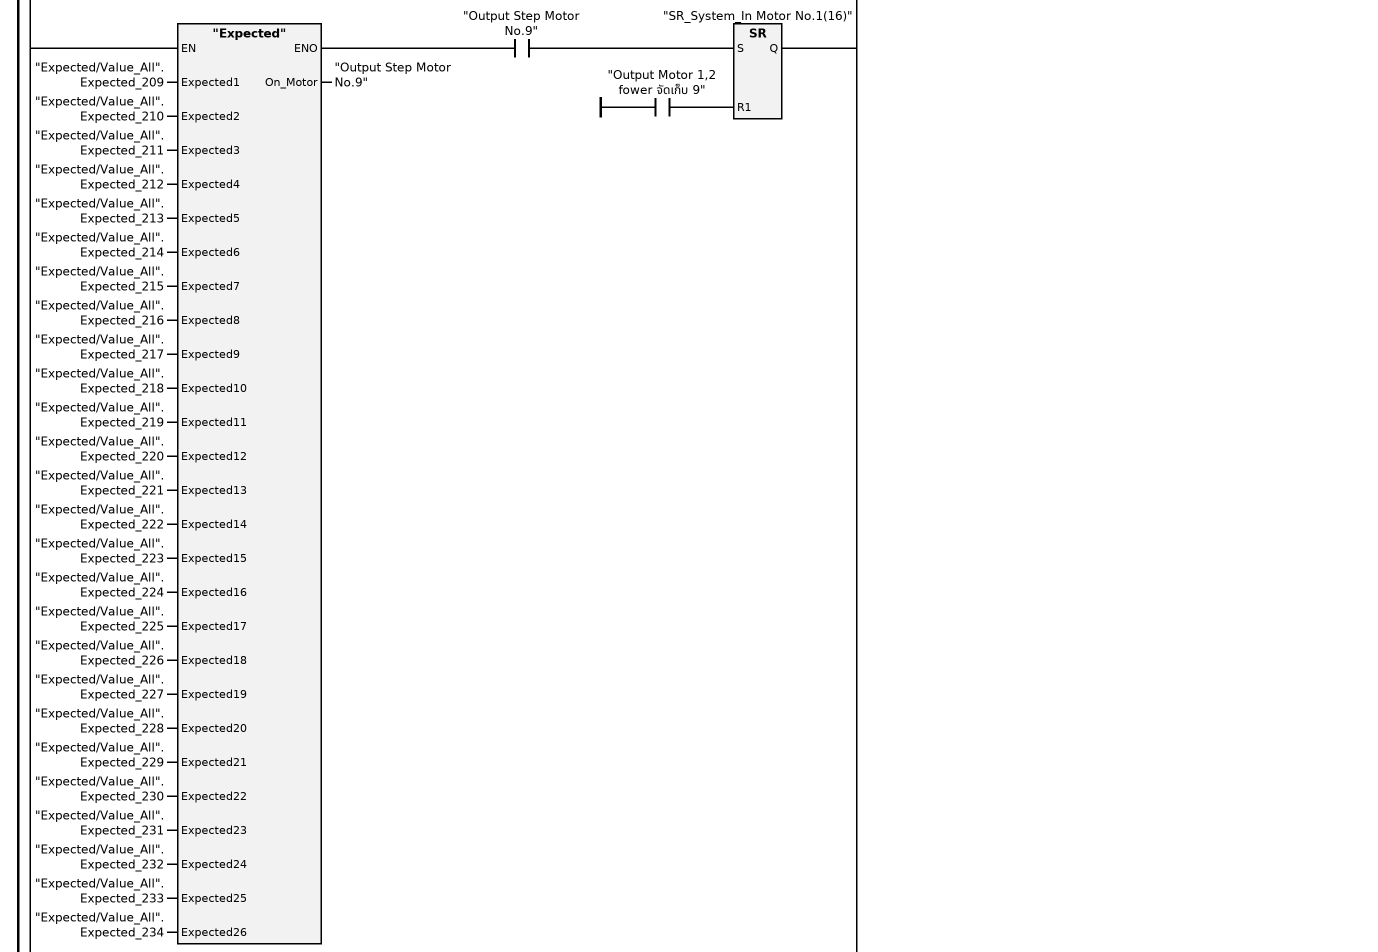
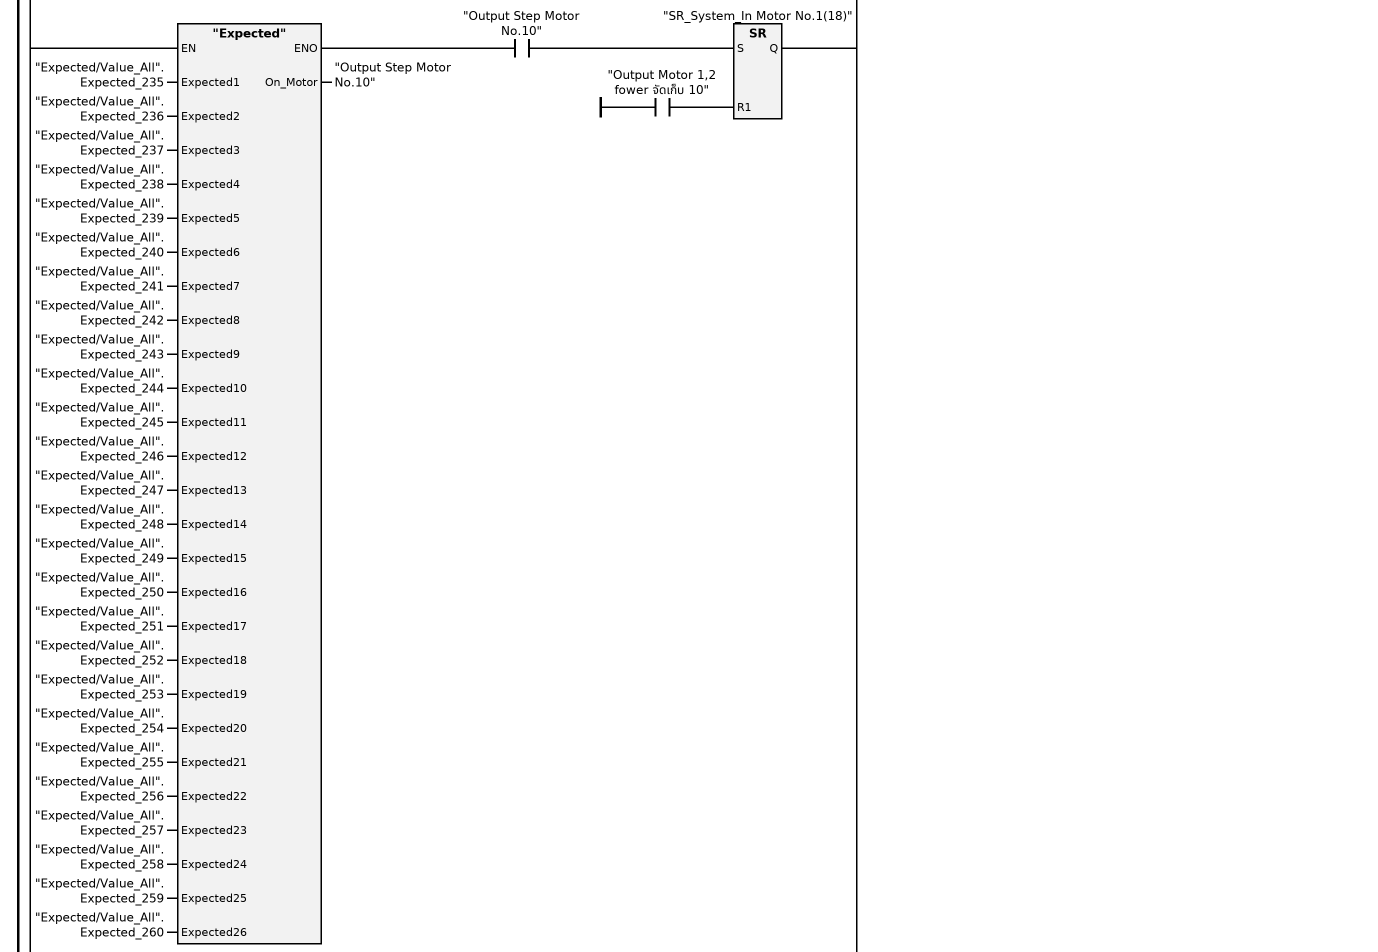
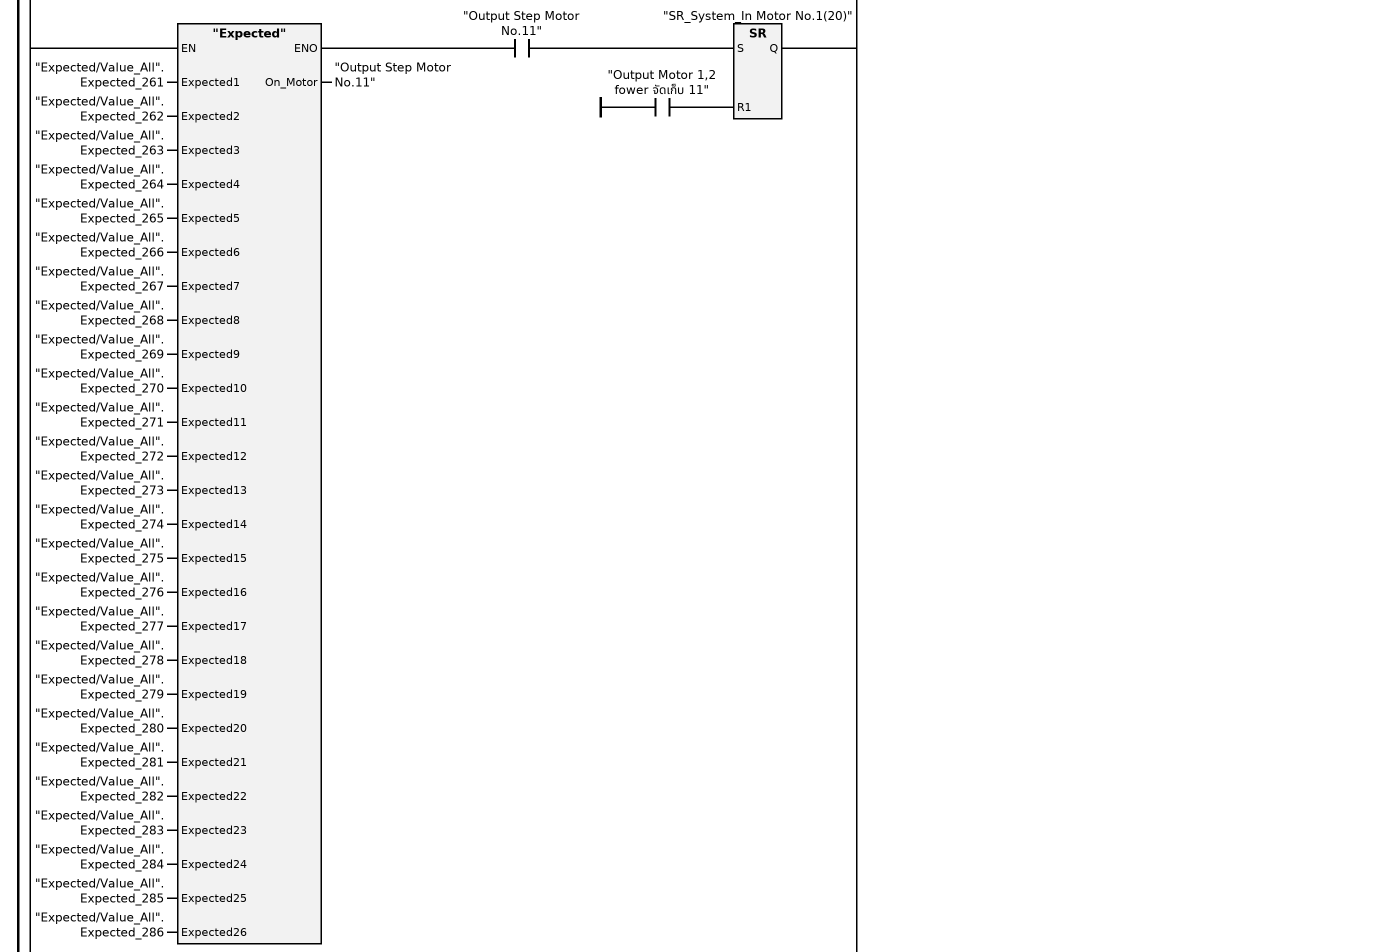
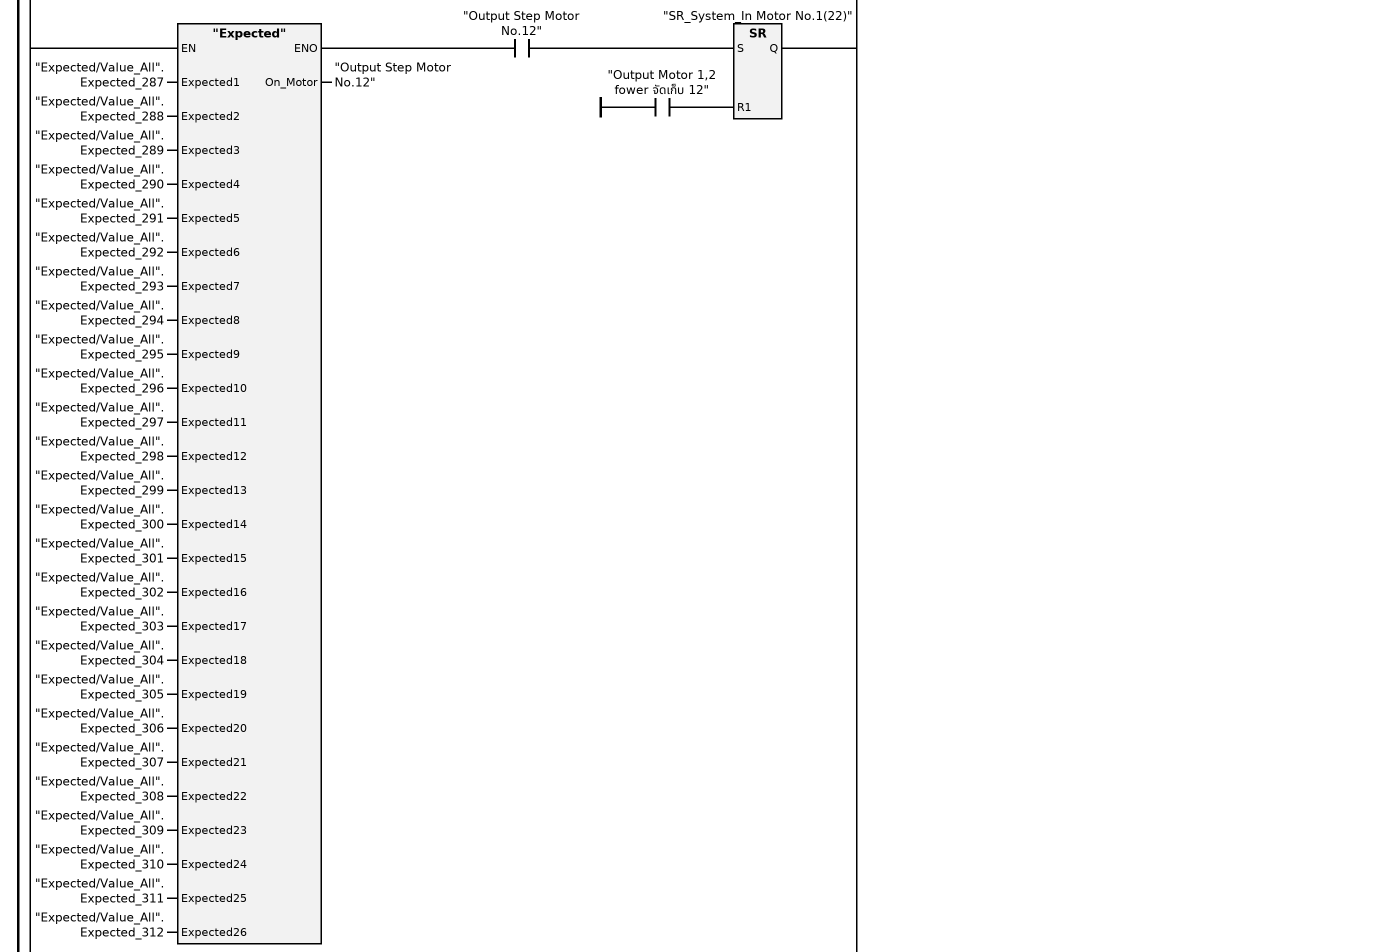
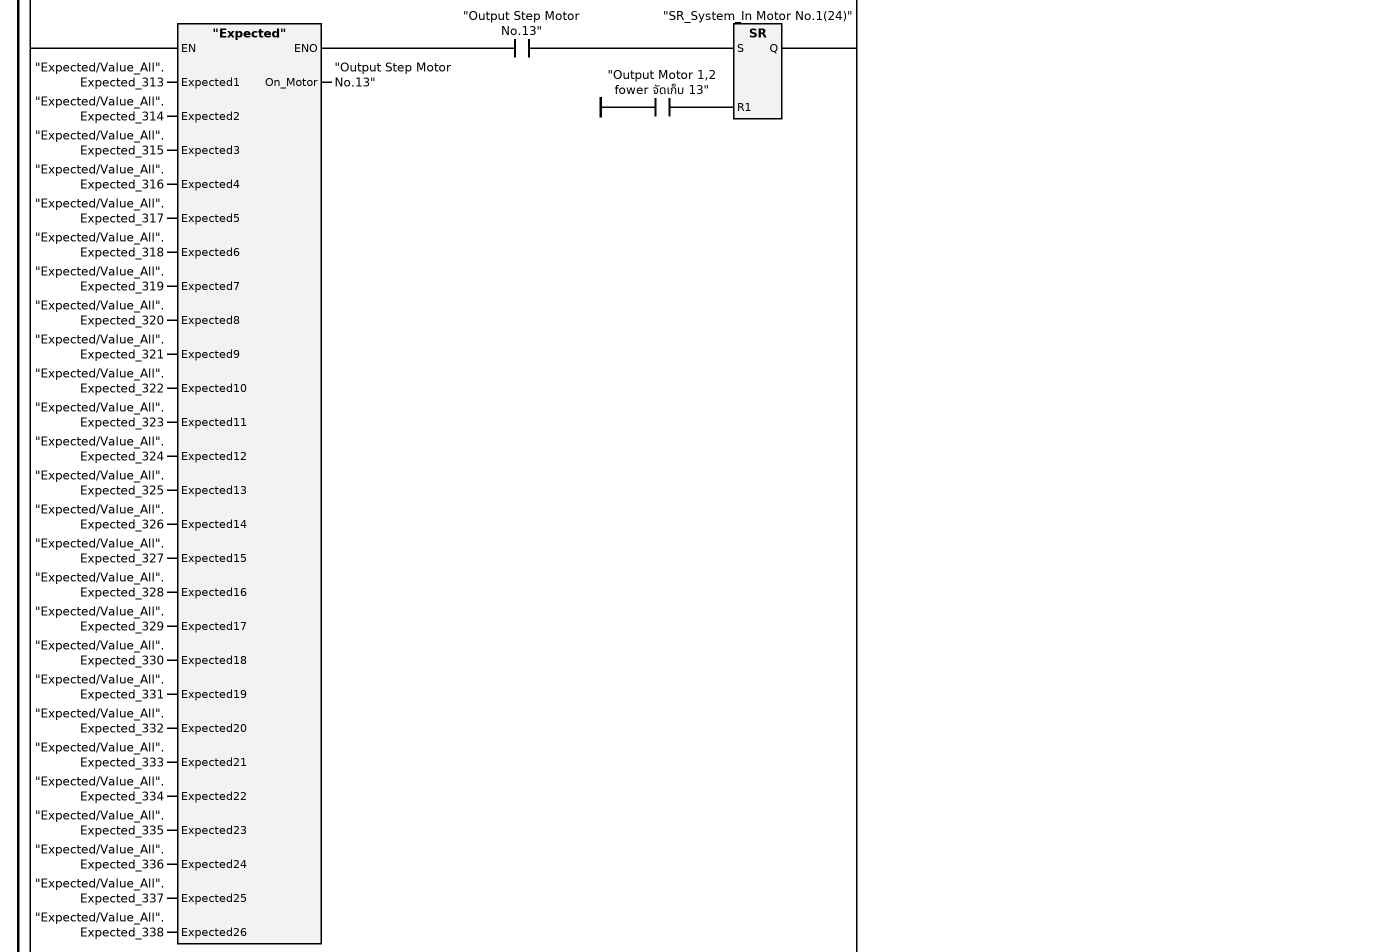
